(* IEC 61131-3 sources: stf-hw/web/public/sil (part 2) *)

(* HBW belt and the two RFID read points. Generated by stf-cad/hbw/sil/iec.py from the proven motion (control.py); do not edit. *)
FUNCTION_BLOCK FB_Belt
VAR_INPUT
    Enable : BOOL;        (* K0 safety relay OK AND mode = AUTO *)
    Ack : BOOL;           (* HMI acknowledge *)
    Reset : BOOL;         (* S3 reset, via the safety relay *)
    Cmd : INT;            (* job to start (0 = none), taken when READY *)
    Arg1 : INT;           (* binding: slot / bay / slot pair index *)
    I2 : BOOL;           (* phototransistor inside *)
    I3 : BOOL;           (* phototransistor outside *)
    Tag : INT;            (* the mould the record expects at RP2 *)
    ExpI2, ExpI3 : BOOL;  (* the belt's occupancy the record expects *)
    RF1_Valid, RF2_Valid : BOOL;
    RF2_Tag : INT;
END_VAR
VAR_OUTPUT
    Q1 : BOOL;           (* conveyor belt forward (M1) *)
    Q2 : BOOL;           (* conveyor belt backward (M1) *)
    Ready, Busy, Done, Fault : BOOL;   (* Done: one scan, when a job ends *)
    Alarm : INT;          (* the state whose watchdog tripped *)
    Sn : INT;             (* the active state *)
END_VAR
VAR
    Prev : INT := -1;
    Job, B1 : INT;
    Wd : TON;             (* step watchdog *)
    Tm : TON;             (* step timer *)
    WdTime : TIME;        (* the active state's watchdog; 0 = none *)
    RfSeen : BOOL;
END_VAR

(* every scan: outputs off unless the active state sets them; Done is a pulse *)
Q1 := FALSE; Q2 := FALSE; Done := FALSE;
IF NOT Enable AND Sn <> 900 THEN Sn := 900; END_IF;
Wd(IN := (Sn = Prev) AND (WdTime > T#0MS), PT := WdTime);
Tm(IN := (Sn = Prev), PT := T#1H);
IF Sn <> Prev THEN RfSeen := FALSE; END_IF;
RfSeen := RfSeen OR RF1_Valid;
Prev := Sn;
IF Wd.Q THEN Alarm := Sn; Sn := 910; END_IF;

CASE Sn OF
  0: (* INIT: power-up, all outputs off *)
      WdTime := T#0MS; IF Enable THEN Sn := 10; END_IF;
  10: (* H:check: occupancy check: I2/I3 against the record *)
      WdTime := T#0MS;
      IF (I2 = ExpI2) AND (I3 = ExpI3) THEN Sn := 100; END_IF;
  100: (* READY: homed, waiting for a job *)
      WdTime := T#0MS; Ready := TRUE; Busy := FALSE;
      IF Cmd <> 0 THEN Job := Cmd; B1 := Arg1; Busy := TRUE; Ready := FALSE;
          CASE Cmd OF 10: Sn := 1000; 12: Sn := 2000; ELSE Sn := 910; Alarm := -Cmd; END_CASE;
      END_IF;
  1000: (* belt_back.01 RP2: RP2 reads the tag of the mould going in *)
      WdTime := T#900MS;
      IF RF2_Valid AND RF2_Tag = Tag THEN Sn := 1001; END_IF;
  1001: (* belt_back.02 run->I2: belt back to the crane; RP1 reads the tag on the fly *)
      WdTime := T#8100MS;
      Q2 := TRUE;
      IF I2 AND RfSeen THEN Done := TRUE; Busy := FALSE; Sn := 100; END_IF;
  2000: (* belt_fwd.01 run->I3: belt out to the VGR hand-over; RP1 reads the tag on the fly *)
      WdTime := T#8100MS;
      Q1 := TRUE;
      IF I3 AND RfSeen THEN Sn := 2001; END_IF;
  2001: (* belt_fwd.02 RP2: RP2 reads the tag at rest and compares it with the record *)
      WdTime := T#900MS;
      IF RF2_Valid AND RF2_Tag = Tag THEN Done := TRUE; Busy := FALSE; Sn := 100; END_IF;
  900: (* ESTOP: the safety relay dropped, outputs off *)
      WdTime := T#0MS; Busy := FALSE; Ready := FALSE; IF Reset AND Enable THEN Sn := 0; END_IF;
  910: (* FAULT: a step timed out, outputs off, alarm raised *)
      WdTime := T#0MS; Fault := TRUE; Busy := FALSE; Ready := FALSE;
      IF Ack AND Enable THEN Fault := FALSE; Sn := 10; END_IF;
END_CASE;
END_FUNCTION_BLOCK

(* VGR arm and vacuum. Generated by stf-cad/hbw/sil/iec.py from the proven motion (control.py); do not edit. *)
FUNCTION_BLOCK FB_Arm
VAR_INPUT
    Enable : BOOL;        (* K0 safety relay OK AND mode = AUTO *)
    Ack : BOOL;           (* HMI acknowledge *)
    Reset : BOOL;         (* S3 reset, via the safety relay *)
    Cmd : INT;            (* job to start (0 = none), taken when READY *)
    Arg1 : INT;           (* binding: slot / bay / slot pair index *)
    I1 : BOOL;           (* reference vertical *)
    I2 : BOOL;           (* reference horizontal *)
    I3 : BOOL;           (* reference rotate *)
    I4 : BOOL;           (* vacuum switch: the cup is sealed on a part (-0.3 bar) *)
    PosPlunge : REAL;     (* plunge, from the encoder counter *)
    PosReach : REAL;     (* reach, from the encoder counter *)
    PosSwivel : REAL;     (* swivel, from the encoder counter *)
END_VAR
VAR_OUTPUT
    Q1 : BOOL;           (* vertical up (M1) *)
    Q2 : BOOL;           (* vertical down (M1) *)
    Q3 : BOOL;           (* horizontal backward (M2) *)
    Q4 : BOOL;           (* horizontal forward (M2) *)
    Q5 : BOOL;           (* rotate clockwise (M3) *)
    Q6 : BOOL;           (* rotate counter-clockwise (M3) *)
    Q8 : BOOL;           (*  *)
    Ready, Busy, Done, Fault : BOOL;   (* Done: one scan, when a job ends *)
    Alarm : INT;          (* the state whose watchdog tripped *)
    Sn : INT;             (* the active state *)
END_VAR
VAR
    Prev : INT := -1;
    Job, B1 : INT;
    Wd : TON;             (* step watchdog *)
    Tm : TON;             (* step timer *)
    WdTime : TIME;        (* the active state's watchdog; 0 = none *)
END_VAR
VAR CONSTANT
    TG_PLACE_OVEN_PLUNGE : ARRAY[1..1, 1..11] OF REAL := [240.0, 153.0, 153.0, 108.0, 104.0, 0.0, 108.0, 153.0, 153.0, 500.0, 500.0];
    TG_PLACE_OVEN_REACH : ARRAY[1..1, 1..11] OF REAL := [301.376, 365.895, 365.895, 365.895, 365.895, 0.0, 365.895, 365.895, 365.895, 0.0, 0.0];
    TG_PLACE_OVEN_SWIVEL : ARRAY[1..1, 1..11] OF REAL := [46.205, 23.396, 23.396, 23.396, 23.396, 0.0, 23.396, 23.396, 23.396, 0.0, 0.0];
    TG_BELT_TO_OVEN_PLUNGE : ARRAY[1..1, 1..10] OF REAL := [500.0, 201.0, 201.0, 156.0, 152.0, 0.0, 156.0, 201.0, 201.0, 240.0];
    TG_BELT_TO_OVEN_REACH : ARRAY[1..1, 1..10] OF REAL := [0.0, 236.857, 236.857, 236.857, 236.857, 0.0, 236.857, 236.857, 236.857, 301.376];
    TG_BELT_TO_OVEN_SWIVEL : ARRAY[1..1, 1..10] OF REAL := [0.0, 69.013, 69.013, 69.013, 69.013, 0.0, 69.013, 69.013, 69.013, 46.205];
    TG_BAY_TO_BELT_PLUNGE : ARRAY[1..3, 1..21] OF REAL := [500.0, 138.0, 138.0, 93.0, 89.0, 0.0, 93.0, 138.0, 138.0, 240.0, 240.0, 201.0, 201.0, 156.0, 152.0, 0.0, 156.0, 201.0, 201.0, 500.0, 500.0, 500.0, 138.0, 138.0, 93.0, 89.0, 0.0, 93.0, 138.0, 138.0, 240.0, 240.0, 201.0, 201.0, 156.0, 152.0, 0.0, 156.0, 201.0, 201.0, 500.0, 500.0, 500.0, 138.0, 138.0, 93.0, 89.0, 0.0, 93.0, 138.0, 138.0, 240.0, 240.0, 201.0, 201.0, 156.0, 152.0, 0.0, 156.0, 201.0, 201.0, 500.0, 500.0];
    TG_BAY_TO_BELT_REACH : ARRAY[1..3, 1..21] OF REAL := [0.0, 157.983, 157.983, 157.983, 157.983, 0.0, 157.983, 157.983, 157.983, 197.42, 197.42, 236.857, 236.857, 236.857, 236.857, 0.0, 236.857, 236.857, 236.857, 0.0, 0.0, 0.0, 155.396, 155.396, 155.396, 155.396, 0.0, 155.396, 155.396, 155.396, 196.126, 196.126, 236.857, 236.857, 236.857, 236.857, 0.0, 236.857, 236.857, 236.857, 0.0, 0.0, 0.0, 208.968, 208.968, 208.968, 208.968, 0.0, 208.968, 208.968, 208.968, 222.912, 222.912, 236.857, 236.857, 236.857, 236.857, 0.0, 236.857, 236.857, 236.857, 0.0, 0.0];
    TG_BAY_TO_BELT_SWIVEL : ARRAY[1..3, 1..21] OF REAL := [0.0, -76.518, -76.518, -76.518, -76.518, 0.0, -76.518, -76.518, -76.518, -3.752, -3.752, 69.013, 69.013, 69.013, 69.013, 0.0, 69.013, 69.013, 69.013, 0.0, 0.0, 0.0, -101.414, -101.414, -101.414, -101.414, 0.0, -101.414, -101.414, -101.414, -16.2, -16.2, 69.013, 69.013, 69.013, 69.013, 0.0, 69.013, 69.013, 69.013, 0.0, 0.0, 0.0, -122.763, -122.763, -122.763, -122.763, 0.0, -122.763, -122.763, -122.763, -26.875, -26.875, 69.013, 69.013, 69.013, 69.013, 0.0, 69.013, 69.013, 69.013, 0.0, 0.0];
    WD_BAY_TO_BELT : ARRAY[1..3, 1..21] OF TIME := [T#600MS, T#5000MS, T#600MS, T#1100MS, T#1100MS, T#1200MS, T#1100MS, T#1100MS, T#600MS, T#2300MS, T#600MS, T#2300MS, T#600MS, T#1100MS, T#1100MS, T#900MS, T#1100MS, T#1100MS, T#600MS, T#4200MS, T#600MS, T#600MS, T#5000MS, T#600MS, T#1100MS, T#1100MS, T#1200MS, T#1100MS, T#1100MS, T#600MS, T#2600MS, T#600MS, T#2600MS, T#600MS, T#1100MS, T#1100MS, T#900MS, T#1100MS, T#1100MS, T#600MS, T#4200MS, T#600MS, T#600MS, T#5000MS, T#600MS, T#1100MS, T#1100MS, T#1200MS, T#1100MS, T#1100MS, T#600MS, T#2900MS, T#600MS, T#2900MS, T#600MS, T#1100MS, T#1100MS, T#900MS, T#1100MS, T#1100MS, T#600MS, T#4200MS, T#600MS];
END_VAR

(* every scan: outputs off unless the active state sets them; Done is a pulse *)
Q1 := FALSE; Q2 := FALSE; Q3 := FALSE; Q4 := FALSE; Q5 := FALSE; Q6 := FALSE; Q8 := FALSE; Done := FALSE;
IF NOT Enable AND Sn <> 900 THEN Sn := 900; END_IF;
Wd(IN := (Sn = Prev) AND (WdTime > T#0MS), PT := WdTime);
Tm(IN := (Sn = Prev), PT := T#1H);
Prev := Sn;
IF Wd.Q THEN Alarm := Sn; Sn := 910; END_IF;

CASE Sn OF
  0: (* INIT: power-up, all outputs off *)
      WdTime := T#0MS; IF Enable THEN Sn := 10; END_IF;
  10: (* H:plunge: plunge up to the reference switch *)
      WdTime := T#6200MS;
      Q1 := TRUE;
      IF I1 THEN Sn := 11; END_IF;
  11: (* H:reach: reach back to the reference switch *)
      WdTime := T#5500MS;
      Q3 := TRUE;
      IF I2 THEN Sn := 12; END_IF;
  12: (* H:swivel: swivel to the reference switch *)
      WdTime := T#7000MS;
      Q6 := TRUE;
      IF I3 THEN Sn := 100; END_IF;
  100: (* READY: homed, waiting for a job *)
      WdTime := T#0MS; Ready := TRUE; Busy := FALSE;
      IF Cmd <> 0 THEN Job := Cmd; B1 := Arg1; Busy := TRUE; Ready := FALSE;
          CASE Cmd OF 7: Sn := 1000; 8: Sn := 2000; 9: Sn := 3000; ELSE Sn := 910; Alarm := -Cmd; END_CASE;
      END_IF;
  1000: (* place_oven.01 k11:pos: swing to the target at transit height *)
      WdTime := T#600MS;
      Q8 := TRUE;
      CASE Drive(PosPlunge, TG_PLACE_OVEN_PLUNGE[B1, 1], 0.3) OF -1: Q2 := TRUE; 1: Q1 := TRUE; END_CASE;
      CASE Drive(PosReach, TG_PLACE_OVEN_REACH[B1, 1], 0.3) OF -1: Q3 := TRUE; 1: Q4 := TRUE; END_CASE;
      CASE Drive(PosSwivel, TG_PLACE_OVEN_SWIVEL[B1, 1], 0.15) OF -1: Q6 := TRUE; 1: Q5 := TRUE; END_CASE;
      IF ABS(PosPlunge - TG_PLACE_OVEN_PLUNGE[B1, 1]) <= 4.0 AND ABS(PosReach - TG_PLACE_OVEN_REACH[B1, 1]) <= 2.5 AND ABS(PosSwivel - TG_PLACE_OVEN_SWIVEL[B1, 1]) <= 0.252 THEN Sn := 1001; END_IF;
  1001: (* place_oven.02 k12:pos: descend beside the target *)
      WdTime := T#1600MS;
      Q8 := TRUE;
      CASE Drive(PosPlunge, TG_PLACE_OVEN_PLUNGE[B1, 2], 0.3) OF -1: Q2 := TRUE; 1: Q1 := TRUE; END_CASE;
      CASE Drive(PosReach, TG_PLACE_OVEN_REACH[B1, 2], 0.3) OF -1: Q3 := TRUE; 1: Q4 := TRUE; END_CASE;
      CASE Drive(PosSwivel, TG_PLACE_OVEN_SWIVEL[B1, 2], 0.15) OF -1: Q6 := TRUE; 1: Q5 := TRUE; END_CASE;
      IF ABS(PosPlunge - TG_PLACE_OVEN_PLUNGE[B1, 2]) <= 4.0 AND ABS(PosReach - TG_PLACE_OVEN_REACH[B1, 2]) <= 2.5 AND ABS(PosSwivel - TG_PLACE_OVEN_SWIVEL[B1, 2]) <= 0.252 THEN Sn := 1002; END_IF;
  1002: (* place_oven.03 k13:pos: extend over the target *)
      WdTime := T#600MS;
      Q8 := TRUE;
      CASE Drive(PosPlunge, TG_PLACE_OVEN_PLUNGE[B1, 3], 0.3) OF -1: Q2 := TRUE; 1: Q1 := TRUE; END_CASE;
      CASE Drive(PosReach, TG_PLACE_OVEN_REACH[B1, 3], 0.3) OF -1: Q3 := TRUE; 1: Q4 := TRUE; END_CASE;
      CASE Drive(PosSwivel, TG_PLACE_OVEN_SWIVEL[B1, 3], 0.15) OF -1: Q6 := TRUE; 1: Q5 := TRUE; END_CASE;
      IF ABS(PosPlunge - TG_PLACE_OVEN_PLUNGE[B1, 3]) <= 4.0 AND ABS(PosReach - TG_PLACE_OVEN_REACH[B1, 3]) <= 2.5 AND ABS(PosSwivel - TG_PLACE_OVEN_SWIVEL[B1, 3]) <= 0.252 THEN Sn := 1003; END_IF;
  1003: (* place_oven.04 k14:pos: cup meets the cookie's top face *)
      WdTime := T#1100MS;
      Q8 := TRUE;
      CASE Drive(PosPlunge, TG_PLACE_OVEN_PLUNGE[B1, 4], 0.3) OF -1: Q2 := TRUE; 1: Q1 := TRUE; END_CASE;
      CASE Drive(PosReach, TG_PLACE_OVEN_REACH[B1, 4], 0.3) OF -1: Q3 := TRUE; 1: Q4 := TRUE; END_CASE;
      CASE Drive(PosSwivel, TG_PLACE_OVEN_SWIVEL[B1, 4], 0.15) OF -1: Q6 := TRUE; 1: Q5 := TRUE; END_CASE;
      IF ABS(PosPlunge - TG_PLACE_OVEN_PLUNGE[B1, 4]) <= 4.0 AND ABS(PosReach - TG_PLACE_OVEN_REACH[B1, 4]) <= 2.5 AND ABS(PosSwivel - TG_PLACE_OVEN_SWIVEL[B1, 4]) <= 0.252 THEN Sn := 1004; END_IF;
  1004: (* place_oven.05 k15:pos: press: the spring stem takes up the over-travel *)
      WdTime := T#1100MS;
      Q8 := TRUE;
      CASE Drive(PosPlunge, TG_PLACE_OVEN_PLUNGE[B1, 5], 0.3) OF -1: Q2 := TRUE; 1: Q1 := TRUE; END_CASE;
      CASE Drive(PosReach, TG_PLACE_OVEN_REACH[B1, 5], 0.3) OF -1: Q3 := TRUE; 1: Q4 := TRUE; END_CASE;
      CASE Drive(PosSwivel, TG_PLACE_OVEN_SWIVEL[B1, 5], 0.15) OF -1: Q6 := TRUE; 1: Q5 := TRUE; END_CASE;
      IF ABS(PosPlunge - TG_PLACE_OVEN_PLUNGE[B1, 5]) <= 4.0 AND ABS(PosReach - TG_PLACE_OVEN_REACH[B1, 5]) <= 2.5 AND ABS(PosSwivel - TG_PLACE_OVEN_SWIVEL[B1, 5]) <= 0.252 THEN Sn := 1005; END_IF;
  1005: (* place_oven.06 k16:vac: Q8 off: the cookie is released (I4 drops) *)
      WdTime := T#900MS;
      IF NOT I4 THEN Sn := 1006; END_IF;
  1006: (* place_oven.07 k17:pos: spring relaxes *)
      WdTime := T#1100MS;
      CASE Drive(PosPlunge, TG_PLACE_OVEN_PLUNGE[B1, 7], 0.3) OF -1: Q2 := TRUE; 1: Q1 := TRUE; END_CASE;
      CASE Drive(PosReach, TG_PLACE_OVEN_REACH[B1, 7], 0.3) OF -1: Q3 := TRUE; 1: Q4 := TRUE; END_CASE;
      CASE Drive(PosSwivel, TG_PLACE_OVEN_SWIVEL[B1, 7], 0.15) OF -1: Q6 := TRUE; 1: Q5 := TRUE; END_CASE;
      IF ABS(PosPlunge - TG_PLACE_OVEN_PLUNGE[B1, 7]) <= 4.0 AND ABS(PosReach - TG_PLACE_OVEN_REACH[B1, 7]) <= 2.5 AND ABS(PosSwivel - TG_PLACE_OVEN_SWIVEL[B1, 7]) <= 0.252 THEN Sn := 1007; END_IF;
  1007: (* place_oven.08 k18:pos: lift clear *)
      WdTime := T#1100MS;
      CASE Drive(PosPlunge, TG_PLACE_OVEN_PLUNGE[B1, 8], 0.3) OF -1: Q2 := TRUE; 1: Q1 := TRUE; END_CASE;
      CASE Drive(PosReach, TG_PLACE_OVEN_REACH[B1, 8], 0.3) OF -1: Q3 := TRUE; 1: Q4 := TRUE; END_CASE;
      CASE Drive(PosSwivel, TG_PLACE_OVEN_SWIVEL[B1, 8], 0.15) OF -1: Q6 := TRUE; 1: Q5 := TRUE; END_CASE;
      IF ABS(PosPlunge - TG_PLACE_OVEN_PLUNGE[B1, 8]) <= 4.0 AND ABS(PosReach - TG_PLACE_OVEN_REACH[B1, 8]) <= 2.5 AND ABS(PosSwivel - TG_PLACE_OVEN_SWIVEL[B1, 8]) <= 0.252 THEN Sn := 1008; END_IF;
  1008: (* place_oven.09 k19:pos: retract out from the station *)
      WdTime := T#600MS;
      CASE Drive(PosPlunge, TG_PLACE_OVEN_PLUNGE[B1, 9], 0.3) OF -1: Q2 := TRUE; 1: Q1 := TRUE; END_CASE;
      CASE Drive(PosReach, TG_PLACE_OVEN_REACH[B1, 9], 0.3) OF -1: Q3 := TRUE; 1: Q4 := TRUE; END_CASE;
      CASE Drive(PosSwivel, TG_PLACE_OVEN_SWIVEL[B1, 9], 0.15) OF -1: Q6 := TRUE; 1: Q5 := TRUE; END_CASE;
      IF ABS(PosPlunge - TG_PLACE_OVEN_PLUNGE[B1, 9]) <= 4.0 AND ABS(PosReach - TG_PLACE_OVEN_REACH[B1, 9]) <= 2.5 AND ABS(PosSwivel - TG_PLACE_OVEN_SWIVEL[B1, 9]) <= 0.252 THEN Sn := 1009; END_IF;
  1009: (* place_oven.10 k20:pos: rise to transit height *)
      WdTime := T#5100MS;
      CASE Drive(PosPlunge, TG_PLACE_OVEN_PLUNGE[B1, 10], 0.3) OF -1: Q2 := TRUE; 1: Q1 := TRUE; END_CASE;
      CASE Drive(PosReach, TG_PLACE_OVEN_REACH[B1, 10], 0.3) OF -1: Q3 := TRUE; 1: Q4 := TRUE; END_CASE;
      CASE Drive(PosSwivel, TG_PLACE_OVEN_SWIVEL[B1, 10], 0.15) OF -1: Q6 := TRUE; 1: Q5 := TRUE; END_CASE;
      IF ABS(PosPlunge - TG_PLACE_OVEN_PLUNGE[B1, 10]) <= 4.0 AND ABS(PosReach - TG_PLACE_OVEN_REACH[B1, 10]) <= 2.5 AND ABS(PosSwivel - TG_PLACE_OVEN_SWIVEL[B1, 10]) <= 0.252 THEN Sn := 1010; END_IF;
  1010: (* place_oven.11 k21:pos: VGR back home *)
      WdTime := T#600MS;
      CASE Drive(PosPlunge, TG_PLACE_OVEN_PLUNGE[B1, 11], 0.3) OF -1: Q2 := TRUE; 1: Q1 := TRUE; END_CASE;
      CASE Drive(PosReach, TG_PLACE_OVEN_REACH[B1, 11], 0.3) OF -1: Q3 := TRUE; 1: Q4 := TRUE; END_CASE;
      CASE Drive(PosSwivel, TG_PLACE_OVEN_SWIVEL[B1, 11], 0.15) OF -1: Q6 := TRUE; 1: Q5 := TRUE; END_CASE;
      IF ABS(PosPlunge - TG_PLACE_OVEN_PLUNGE[B1, 11]) <= 4.0 AND ABS(PosReach - TG_PLACE_OVEN_REACH[B1, 11]) <= 2.5 AND ABS(PosSwivel - TG_PLACE_OVEN_SWIVEL[B1, 11]) <= 0.252 THEN Done := TRUE; Busy := FALSE; Sn := 100; END_IF;
  2000: (* belt_to_oven.01 k1:pos: swing to the source at transit height *)
      WdTime := T#600MS;
      CASE Drive(PosPlunge, TG_BELT_TO_OVEN_PLUNGE[B1, 1], 0.3) OF -1: Q2 := TRUE; 1: Q1 := TRUE; END_CASE;
      CASE Drive(PosReach, TG_BELT_TO_OVEN_REACH[B1, 1], 0.3) OF -1: Q3 := TRUE; 1: Q4 := TRUE; END_CASE;
      CASE Drive(PosSwivel, TG_BELT_TO_OVEN_SWIVEL[B1, 1], 0.15) OF -1: Q6 := TRUE; 1: Q5 := TRUE; END_CASE;
      IF ABS(PosPlunge - TG_BELT_TO_OVEN_PLUNGE[B1, 1]) <= 4.0 AND ABS(PosReach - TG_BELT_TO_OVEN_REACH[B1, 1]) <= 2.5 AND ABS(PosSwivel - TG_BELT_TO_OVEN_SWIVEL[B1, 1]) <= 0.252 THEN Sn := 2001; END_IF;
  2001: (* belt_to_oven.02 k2:pos: descend beside the source *)
      WdTime := T#4200MS;
      CASE Drive(PosPlunge, TG_BELT_TO_OVEN_PLUNGE[B1, 2], 0.3) OF -1: Q2 := TRUE; 1: Q1 := TRUE; END_CASE;
      CASE Drive(PosReach, TG_BELT_TO_OVEN_REACH[B1, 2], 0.3) OF -1: Q3 := TRUE; 1: Q4 := TRUE; END_CASE;
      CASE Drive(PosSwivel, TG_BELT_TO_OVEN_SWIVEL[B1, 2], 0.15) OF -1: Q6 := TRUE; 1: Q5 := TRUE; END_CASE;
      IF ABS(PosPlunge - TG_BELT_TO_OVEN_PLUNGE[B1, 2]) <= 4.0 AND ABS(PosReach - TG_BELT_TO_OVEN_REACH[B1, 2]) <= 2.5 AND ABS(PosSwivel - TG_BELT_TO_OVEN_SWIVEL[B1, 2]) <= 0.252 THEN Sn := 2002; END_IF;
  2002: (* belt_to_oven.03 k3:pos: extend over the source *)
      WdTime := T#600MS;
      CASE Drive(PosPlunge, TG_BELT_TO_OVEN_PLUNGE[B1, 3], 0.3) OF -1: Q2 := TRUE; 1: Q1 := TRUE; END_CASE;
      CASE Drive(PosReach, TG_BELT_TO_OVEN_REACH[B1, 3], 0.3) OF -1: Q3 := TRUE; 1: Q4 := TRUE; END_CASE;
      CASE Drive(PosSwivel, TG_BELT_TO_OVEN_SWIVEL[B1, 3], 0.15) OF -1: Q6 := TRUE; 1: Q5 := TRUE; END_CASE;
      IF ABS(PosPlunge - TG_BELT_TO_OVEN_PLUNGE[B1, 3]) <= 4.0 AND ABS(PosReach - TG_BELT_TO_OVEN_REACH[B1, 3]) <= 2.5 AND ABS(PosSwivel - TG_BELT_TO_OVEN_SWIVEL[B1, 3]) <= 0.252 THEN Sn := 2003; END_IF;
  2003: (* belt_to_oven.04 k4:pos: cup meets the cookie's top face *)
      WdTime := T#1100MS;
      CASE Drive(PosPlunge, TG_BELT_TO_OVEN_PLUNGE[B1, 4], 0.3) OF -1: Q2 := TRUE; 1: Q1 := TRUE; END_CASE;
      CASE Drive(PosReach, TG_BELT_TO_OVEN_REACH[B1, 4], 0.3) OF -1: Q3 := TRUE; 1: Q4 := TRUE; END_CASE;
      CASE Drive(PosSwivel, TG_BELT_TO_OVEN_SWIVEL[B1, 4], 0.15) OF -1: Q6 := TRUE; 1: Q5 := TRUE; END_CASE;
      IF ABS(PosPlunge - TG_BELT_TO_OVEN_PLUNGE[B1, 4]) <= 4.0 AND ABS(PosReach - TG_BELT_TO_OVEN_REACH[B1, 4]) <= 2.5 AND ABS(PosSwivel - TG_BELT_TO_OVEN_SWIVEL[B1, 4]) <= 0.252 THEN Sn := 2004; END_IF;
  2004: (* belt_to_oven.05 k5:pos: press: the spring stem takes up the over-travel *)
      WdTime := T#1100MS;
      CASE Drive(PosPlunge, TG_BELT_TO_OVEN_PLUNGE[B1, 5], 0.3) OF -1: Q2 := TRUE; 1: Q1 := TRUE; END_CASE;
      CASE Drive(PosReach, TG_BELT_TO_OVEN_REACH[B1, 5], 0.3) OF -1: Q3 := TRUE; 1: Q4 := TRUE; END_CASE;
      CASE Drive(PosSwivel, TG_BELT_TO_OVEN_SWIVEL[B1, 5], 0.15) OF -1: Q6 := TRUE; 1: Q5 := TRUE; END_CASE;
      IF ABS(PosPlunge - TG_BELT_TO_OVEN_PLUNGE[B1, 5]) <= 4.0 AND ABS(PosReach - TG_BELT_TO_OVEN_REACH[B1, 5]) <= 2.5 AND ABS(PosSwivel - TG_BELT_TO_OVEN_SWIVEL[B1, 5]) <= 0.252 THEN Sn := 2005; END_IF;
  2005: (* belt_to_oven.06 k6:vac: Q8 vacuum on: the cup seals on the cookie (I4 made) *)
      WdTime := T#1200MS;
      Q8 := TRUE;
      IF I4 THEN Sn := 2006; END_IF;
  2006: (* belt_to_oven.07 k7:pos: spring relaxes - seal holds *)
      WdTime := T#1100MS;
      Q8 := TRUE;
      CASE Drive(PosPlunge, TG_BELT_TO_OVEN_PLUNGE[B1, 7], 0.3) OF -1: Q2 := TRUE; 1: Q1 := TRUE; END_CASE;
      CASE Drive(PosReach, TG_BELT_TO_OVEN_REACH[B1, 7], 0.3) OF -1: Q3 := TRUE; 1: Q4 := TRUE; END_CASE;
      CASE Drive(PosSwivel, TG_BELT_TO_OVEN_SWIVEL[B1, 7], 0.15) OF -1: Q6 := TRUE; 1: Q5 := TRUE; END_CASE;
      IF ABS(PosPlunge - TG_BELT_TO_OVEN_PLUNGE[B1, 7]) <= 4.0 AND ABS(PosReach - TG_BELT_TO_OVEN_REACH[B1, 7]) <= 2.5 AND ABS(PosSwivel - TG_BELT_TO_OVEN_SWIVEL[B1, 7]) <= 0.252 THEN Sn := 2007; END_IF;
  2007: (* belt_to_oven.08 k8:pos: lift the cookie clear *)
      WdTime := T#1100MS;
      Q8 := TRUE;
      CASE Drive(PosPlunge, TG_BELT_TO_OVEN_PLUNGE[B1, 8], 0.3) OF -1: Q2 := TRUE; 1: Q1 := TRUE; END_CASE;
      CASE Drive(PosReach, TG_BELT_TO_OVEN_REACH[B1, 8], 0.3) OF -1: Q3 := TRUE; 1: Q4 := TRUE; END_CASE;
      CASE Drive(PosSwivel, TG_BELT_TO_OVEN_SWIVEL[B1, 8], 0.15) OF -1: Q6 := TRUE; 1: Q5 := TRUE; END_CASE;
      IF ABS(PosPlunge - TG_BELT_TO_OVEN_PLUNGE[B1, 8]) <= 4.0 AND ABS(PosReach - TG_BELT_TO_OVEN_REACH[B1, 8]) <= 2.5 AND ABS(PosSwivel - TG_BELT_TO_OVEN_SWIVEL[B1, 8]) <= 0.252 THEN Sn := 2008; END_IF;
  2008: (* belt_to_oven.09 k9:pos: retract out from the station *)
      WdTime := T#600MS;
      Q8 := TRUE;
      CASE Drive(PosPlunge, TG_BELT_TO_OVEN_PLUNGE[B1, 9], 0.3) OF -1: Q2 := TRUE; 1: Q1 := TRUE; END_CASE;
      CASE Drive(PosReach, TG_BELT_TO_OVEN_REACH[B1, 9], 0.3) OF -1: Q3 := TRUE; 1: Q4 := TRUE; END_CASE;
      CASE Drive(PosSwivel, TG_BELT_TO_OVEN_SWIVEL[B1, 9], 0.15) OF -1: Q6 := TRUE; 1: Q5 := TRUE; END_CASE;
      IF ABS(PosPlunge - TG_BELT_TO_OVEN_PLUNGE[B1, 9]) <= 4.0 AND ABS(PosReach - TG_BELT_TO_OVEN_REACH[B1, 9]) <= 2.5 AND ABS(PosSwivel - TG_BELT_TO_OVEN_SWIVEL[B1, 9]) <= 0.252 THEN Sn := 2009; END_IF;
  2009: (* belt_to_oven.10 k10:pos: rise to transit height *)
      WdTime := T#1300MS;
      Q8 := TRUE;
      CASE Drive(PosPlunge, TG_BELT_TO_OVEN_PLUNGE[B1, 10], 0.3) OF -1: Q2 := TRUE; 1: Q1 := TRUE; END_CASE;
      CASE Drive(PosReach, TG_BELT_TO_OVEN_REACH[B1, 10], 0.3) OF -1: Q3 := TRUE; 1: Q4 := TRUE; END_CASE;
      CASE Drive(PosSwivel, TG_BELT_TO_OVEN_SWIVEL[B1, 10], 0.15) OF -1: Q6 := TRUE; 1: Q5 := TRUE; END_CASE;
      IF ABS(PosPlunge - TG_BELT_TO_OVEN_PLUNGE[B1, 10]) <= 4.0 AND ABS(PosReach - TG_BELT_TO_OVEN_REACH[B1, 10]) <= 2.5 AND ABS(PosSwivel - TG_BELT_TO_OVEN_SWIVEL[B1, 10]) <= 0.252 THEN Done := TRUE; Busy := FALSE; Sn := 100; END_IF;
  3000: (* bay_to_belt.01 k1:pos: swing to the source at transit height *)
      WdTime := T#600MS;
      CASE Drive(PosPlunge, TG_BAY_TO_BELT_PLUNGE[B1, 1], 0.3) OF -1: Q2 := TRUE; 1: Q1 := TRUE; END_CASE;
      CASE Drive(PosReach, TG_BAY_TO_BELT_REACH[B1, 1], 0.3) OF -1: Q3 := TRUE; 1: Q4 := TRUE; END_CASE;
      CASE Drive(PosSwivel, TG_BAY_TO_BELT_SWIVEL[B1, 1], 0.15) OF -1: Q6 := TRUE; 1: Q5 := TRUE; END_CASE;
      IF ABS(PosPlunge - TG_BAY_TO_BELT_PLUNGE[B1, 1]) <= 4.0 AND ABS(PosReach - TG_BAY_TO_BELT_REACH[B1, 1]) <= 2.5 AND ABS(PosSwivel - TG_BAY_TO_BELT_SWIVEL[B1, 1]) <= 0.252 THEN Sn := 3001; END_IF;
  3001: (* bay_to_belt.02 k2:pos: descend beside the source *)
      WdTime := T#5000MS;
      CASE Drive(PosPlunge, TG_BAY_TO_BELT_PLUNGE[B1, 2], 0.3) OF -1: Q2 := TRUE; 1: Q1 := TRUE; END_CASE;
      CASE Drive(PosReach, TG_BAY_TO_BELT_REACH[B1, 2], 0.3) OF -1: Q3 := TRUE; 1: Q4 := TRUE; END_CASE;
      CASE Drive(PosSwivel, TG_BAY_TO_BELT_SWIVEL[B1, 2], 0.15) OF -1: Q6 := TRUE; 1: Q5 := TRUE; END_CASE;
      IF ABS(PosPlunge - TG_BAY_TO_BELT_PLUNGE[B1, 2]) <= 4.0 AND ABS(PosReach - TG_BAY_TO_BELT_REACH[B1, 2]) <= 2.5 AND ABS(PosSwivel - TG_BAY_TO_BELT_SWIVEL[B1, 2]) <= 0.252 THEN Sn := 3002; END_IF;
  3002: (* bay_to_belt.03 k3:pos: extend over the source *)
      WdTime := T#600MS;
      CASE Drive(PosPlunge, TG_BAY_TO_BELT_PLUNGE[B1, 3], 0.3) OF -1: Q2 := TRUE; 1: Q1 := TRUE; END_CASE;
      CASE Drive(PosReach, TG_BAY_TO_BELT_REACH[B1, 3], 0.3) OF -1: Q3 := TRUE; 1: Q4 := TRUE; END_CASE;
      CASE Drive(PosSwivel, TG_BAY_TO_BELT_SWIVEL[B1, 3], 0.15) OF -1: Q6 := TRUE; 1: Q5 := TRUE; END_CASE;
      IF ABS(PosPlunge - TG_BAY_TO_BELT_PLUNGE[B1, 3]) <= 4.0 AND ABS(PosReach - TG_BAY_TO_BELT_REACH[B1, 3]) <= 2.5 AND ABS(PosSwivel - TG_BAY_TO_BELT_SWIVEL[B1, 3]) <= 0.252 THEN Sn := 3003; END_IF;
  3003: (* bay_to_belt.04 k4:pos: cup meets the cookie's top face *)
      WdTime := T#1100MS;
      CASE Drive(PosPlunge, TG_BAY_TO_BELT_PLUNGE[B1, 4], 0.3) OF -1: Q2 := TRUE; 1: Q1 := TRUE; END_CASE;
      CASE Drive(PosReach, TG_BAY_TO_BELT_REACH[B1, 4], 0.3) OF -1: Q3 := TRUE; 1: Q4 := TRUE; END_CASE;
      CASE Drive(PosSwivel, TG_BAY_TO_BELT_SWIVEL[B1, 4], 0.15) OF -1: Q6 := TRUE; 1: Q5 := TRUE; END_CASE;
      IF ABS(PosPlunge - TG_BAY_TO_BELT_PLUNGE[B1, 4]) <= 4.0 AND ABS(PosReach - TG_BAY_TO_BELT_REACH[B1, 4]) <= 2.5 AND ABS(PosSwivel - TG_BAY_TO_BELT_SWIVEL[B1, 4]) <= 0.252 THEN Sn := 3004; END_IF;
  3004: (* bay_to_belt.05 k5:pos: press: the spring stem takes up the over-travel *)
      WdTime := T#1100MS;
      CASE Drive(PosPlunge, TG_BAY_TO_BELT_PLUNGE[B1, 5], 0.3) OF -1: Q2 := TRUE; 1: Q1 := TRUE; END_CASE;
      CASE Drive(PosReach, TG_BAY_TO_BELT_REACH[B1, 5], 0.3) OF -1: Q3 := TRUE; 1: Q4 := TRUE; END_CASE;
      CASE Drive(PosSwivel, TG_BAY_TO_BELT_SWIVEL[B1, 5], 0.15) OF -1: Q6 := TRUE; 1: Q5 := TRUE; END_CASE;
      IF ABS(PosPlunge - TG_BAY_TO_BELT_PLUNGE[B1, 5]) <= 4.0 AND ABS(PosReach - TG_BAY_TO_BELT_REACH[B1, 5]) <= 2.5 AND ABS(PosSwivel - TG_BAY_TO_BELT_SWIVEL[B1, 5]) <= 0.252 THEN Sn := 3005; END_IF;
  3005: (* bay_to_belt.06 k6:vac: Q8 vacuum on: the cup seals on the cookie (I4 made) *)
      WdTime := T#1200MS;
      Q8 := TRUE;
      IF I4 THEN Sn := 3006; END_IF;
  3006: (* bay_to_belt.07 k7:pos: spring relaxes - seal holds *)
      WdTime := T#1100MS;
      Q8 := TRUE;
      CASE Drive(PosPlunge, TG_BAY_TO_BELT_PLUNGE[B1, 7], 0.3) OF -1: Q2 := TRUE; 1: Q1 := TRUE; END_CASE;
      CASE Drive(PosReach, TG_BAY_TO_BELT_REACH[B1, 7], 0.3) OF -1: Q3 := TRUE; 1: Q4 := TRUE; END_CASE;
      CASE Drive(PosSwivel, TG_BAY_TO_BELT_SWIVEL[B1, 7], 0.15) OF -1: Q6 := TRUE; 1: Q5 := TRUE; END_CASE;
      IF ABS(PosPlunge - TG_BAY_TO_BELT_PLUNGE[B1, 7]) <= 4.0 AND ABS(PosReach - TG_BAY_TO_BELT_REACH[B1, 7]) <= 2.5 AND ABS(PosSwivel - TG_BAY_TO_BELT_SWIVEL[B1, 7]) <= 0.252 THEN Sn := 3007; END_IF;
  3007: (* bay_to_belt.08 k8:pos: lift the cookie clear *)
      WdTime := T#1100MS;
      Q8 := TRUE;
      CASE Drive(PosPlunge, TG_BAY_TO_BELT_PLUNGE[B1, 8], 0.3) OF -1: Q2 := TRUE; 1: Q1 := TRUE; END_CASE;
      CASE Drive(PosReach, TG_BAY_TO_BELT_REACH[B1, 8], 0.3) OF -1: Q3 := TRUE; 1: Q4 := TRUE; END_CASE;
      CASE Drive(PosSwivel, TG_BAY_TO_BELT_SWIVEL[B1, 8], 0.15) OF -1: Q6 := TRUE; 1: Q5 := TRUE; END_CASE;
      IF ABS(PosPlunge - TG_BAY_TO_BELT_PLUNGE[B1, 8]) <= 4.0 AND ABS(PosReach - TG_BAY_TO_BELT_REACH[B1, 8]) <= 2.5 AND ABS(PosSwivel - TG_BAY_TO_BELT_SWIVEL[B1, 8]) <= 0.252 THEN Sn := 3008; END_IF;
  3008: (* bay_to_belt.09 k9:pos: retract out from the station *)
      WdTime := T#600MS;
      Q8 := TRUE;
      CASE Drive(PosPlunge, TG_BAY_TO_BELT_PLUNGE[B1, 9], 0.3) OF -1: Q2 := TRUE; 1: Q1 := TRUE; END_CASE;
      CASE Drive(PosReach, TG_BAY_TO_BELT_REACH[B1, 9], 0.3) OF -1: Q3 := TRUE; 1: Q4 := TRUE; END_CASE;
      CASE Drive(PosSwivel, TG_BAY_TO_BELT_SWIVEL[B1, 9], 0.15) OF -1: Q6 := TRUE; 1: Q5 := TRUE; END_CASE;
      IF ABS(PosPlunge - TG_BAY_TO_BELT_PLUNGE[B1, 9]) <= 4.0 AND ABS(PosReach - TG_BAY_TO_BELT_REACH[B1, 9]) <= 2.5 AND ABS(PosSwivel - TG_BAY_TO_BELT_SWIVEL[B1, 9]) <= 0.252 THEN Sn := 3009; END_IF;
  3009: (* bay_to_belt.10 k10:pos: rise to transit height *)
      WdTime := WD_BAY_TO_BELT[B1, 10];
      Q8 := TRUE;
      CASE Drive(PosPlunge, TG_BAY_TO_BELT_PLUNGE[B1, 10], 0.3) OF -1: Q2 := TRUE; 1: Q1 := TRUE; END_CASE;
      CASE Drive(PosReach, TG_BAY_TO_BELT_REACH[B1, 10], 0.3) OF -1: Q3 := TRUE; 1: Q4 := TRUE; END_CASE;
      CASE Drive(PosSwivel, TG_BAY_TO_BELT_SWIVEL[B1, 10], 0.15) OF -1: Q6 := TRUE; 1: Q5 := TRUE; END_CASE;
      IF ABS(PosPlunge - TG_BAY_TO_BELT_PLUNGE[B1, 10]) <= 4.0 AND ABS(PosReach - TG_BAY_TO_BELT_REACH[B1, 10]) <= 2.5 AND ABS(PosSwivel - TG_BAY_TO_BELT_SWIVEL[B1, 10]) <= 0.252 THEN Sn := 3010; END_IF;
  3010: (* bay_to_belt.11 k11:pos: swing to the target at transit height *)
      WdTime := T#600MS;
      Q8 := TRUE;
      CASE Drive(PosPlunge, TG_BAY_TO_BELT_PLUNGE[B1, 11], 0.3) OF -1: Q2 := TRUE; 1: Q1 := TRUE; END_CASE;
      CASE Drive(PosReach, TG_BAY_TO_BELT_REACH[B1, 11], 0.3) OF -1: Q3 := TRUE; 1: Q4 := TRUE; END_CASE;
      CASE Drive(PosSwivel, TG_BAY_TO_BELT_SWIVEL[B1, 11], 0.15) OF -1: Q6 := TRUE; 1: Q5 := TRUE; END_CASE;
      IF ABS(PosPlunge - TG_BAY_TO_BELT_PLUNGE[B1, 11]) <= 4.0 AND ABS(PosReach - TG_BAY_TO_BELT_REACH[B1, 11]) <= 2.5 AND ABS(PosSwivel - TG_BAY_TO_BELT_SWIVEL[B1, 11]) <= 0.252 THEN Sn := 3011; END_IF;
  3011: (* bay_to_belt.12 k12:pos: descend beside the target *)
      WdTime := WD_BAY_TO_BELT[B1, 12];
      Q8 := TRUE;
      CASE Drive(PosPlunge, TG_BAY_TO_BELT_PLUNGE[B1, 12], 0.3) OF -1: Q2 := TRUE; 1: Q1 := TRUE; END_CASE;
      CASE Drive(PosReach, TG_BAY_TO_BELT_REACH[B1, 12], 0.3) OF -1: Q3 := TRUE; 1: Q4 := TRUE; END_CASE;
      CASE Drive(PosSwivel, TG_BAY_TO_BELT_SWIVEL[B1, 12], 0.15) OF -1: Q6 := TRUE; 1: Q5 := TRUE; END_CASE;
      IF ABS(PosPlunge - TG_BAY_TO_BELT_PLUNGE[B1, 12]) <= 4.0 AND ABS(PosReach - TG_BAY_TO_BELT_REACH[B1, 12]) <= 2.5 AND ABS(PosSwivel - TG_BAY_TO_BELT_SWIVEL[B1, 12]) <= 0.252 THEN Sn := 3012; END_IF;
  3012: (* bay_to_belt.13 k13:pos: extend over the target *)
      WdTime := T#600MS;
      Q8 := TRUE;
      CASE Drive(PosPlunge, TG_BAY_TO_BELT_PLUNGE[B1, 13], 0.3) OF -1: Q2 := TRUE; 1: Q1 := TRUE; END_CASE;
      CASE Drive(PosReach, TG_BAY_TO_BELT_REACH[B1, 13], 0.3) OF -1: Q3 := TRUE; 1: Q4 := TRUE; END_CASE;
      CASE Drive(PosSwivel, TG_BAY_TO_BELT_SWIVEL[B1, 13], 0.15) OF -1: Q6 := TRUE; 1: Q5 := TRUE; END_CASE;
      IF ABS(PosPlunge - TG_BAY_TO_BELT_PLUNGE[B1, 13]) <= 4.0 AND ABS(PosReach - TG_BAY_TO_BELT_REACH[B1, 13]) <= 2.5 AND ABS(PosSwivel - TG_BAY_TO_BELT_SWIVEL[B1, 13]) <= 0.252 THEN Sn := 3013; END_IF;
  3013: (* bay_to_belt.14 k14:pos: cup meets the cookie's top face *)
      WdTime := T#1100MS;
      Q8 := TRUE;
      CASE Drive(PosPlunge, TG_BAY_TO_BELT_PLUNGE[B1, 14], 0.3) OF -1: Q2 := TRUE; 1: Q1 := TRUE; END_CASE;
      CASE Drive(PosReach, TG_BAY_TO_BELT_REACH[B1, 14], 0.3) OF -1: Q3 := TRUE; 1: Q4 := TRUE; END_CASE;
      CASE Drive(PosSwivel, TG_BAY_TO_BELT_SWIVEL[B1, 14], 0.15) OF -1: Q6 := TRUE; 1: Q5 := TRUE; END_CASE;
      IF ABS(PosPlunge - TG_BAY_TO_BELT_PLUNGE[B1, 14]) <= 4.0 AND ABS(PosReach - TG_BAY_TO_BELT_REACH[B1, 14]) <= 2.5 AND ABS(PosSwivel - TG_BAY_TO_BELT_SWIVEL[B1, 14]) <= 0.252 THEN Sn := 3014; END_IF;
  3014: (* bay_to_belt.15 k15:pos: press: the spring stem takes up the over-travel *)
      WdTime := T#1100MS;
      Q8 := TRUE;
      CASE Drive(PosPlunge, TG_BAY_TO_BELT_PLUNGE[B1, 15], 0.3) OF -1: Q2 := TRUE; 1: Q1 := TRUE; END_CASE;
      CASE Drive(PosReach, TG_BAY_TO_BELT_REACH[B1, 15], 0.3) OF -1: Q3 := TRUE; 1: Q4 := TRUE; END_CASE;
      CASE Drive(PosSwivel, TG_BAY_TO_BELT_SWIVEL[B1, 15], 0.15) OF -1: Q6 := TRUE; 1: Q5 := TRUE; END_CASE;
      IF ABS(PosPlunge - TG_BAY_TO_BELT_PLUNGE[B1, 15]) <= 4.0 AND ABS(PosReach - TG_BAY_TO_BELT_REACH[B1, 15]) <= 2.5 AND ABS(PosSwivel - TG_BAY_TO_BELT_SWIVEL[B1, 15]) <= 0.252 THEN Sn := 3015; END_IF;
  3015: (* bay_to_belt.16 k16:vac: Q8 off: the cookie is released (I4 drops) *)
      WdTime := T#900MS;
      IF NOT I4 THEN Sn := 3016; END_IF;
  3016: (* bay_to_belt.17 k17:pos: spring relaxes *)
      WdTime := T#1100MS;
      CASE Drive(PosPlunge, TG_BAY_TO_BELT_PLUNGE[B1, 17], 0.3) OF -1: Q2 := TRUE; 1: Q1 := TRUE; END_CASE;
      CASE Drive(PosReach, TG_BAY_TO_BELT_REACH[B1, 17], 0.3) OF -1: Q3 := TRUE; 1: Q4 := TRUE; END_CASE;
      CASE Drive(PosSwivel, TG_BAY_TO_BELT_SWIVEL[B1, 17], 0.15) OF -1: Q6 := TRUE; 1: Q5 := TRUE; END_CASE;
      IF ABS(PosPlunge - TG_BAY_TO_BELT_PLUNGE[B1, 17]) <= 4.0 AND ABS(PosReach - TG_BAY_TO_BELT_REACH[B1, 17]) <= 2.5 AND ABS(PosSwivel - TG_BAY_TO_BELT_SWIVEL[B1, 17]) <= 0.252 THEN Sn := 3017; END_IF;
  3017: (* bay_to_belt.18 k18:pos: lift clear *)
      WdTime := T#1100MS;
      CASE Drive(PosPlunge, TG_BAY_TO_BELT_PLUNGE[B1, 18], 0.3) OF -1: Q2 := TRUE; 1: Q1 := TRUE; END_CASE;
      CASE Drive(PosReach, TG_BAY_TO_BELT_REACH[B1, 18], 0.3) OF -1: Q3 := TRUE; 1: Q4 := TRUE; END_CASE;
      CASE Drive(PosSwivel, TG_BAY_TO_BELT_SWIVEL[B1, 18], 0.15) OF -1: Q6 := TRUE; 1: Q5 := TRUE; END_CASE;
      IF ABS(PosPlunge - TG_BAY_TO_BELT_PLUNGE[B1, 18]) <= 4.0 AND ABS(PosReach - TG_BAY_TO_BELT_REACH[B1, 18]) <= 2.5 AND ABS(PosSwivel - TG_BAY_TO_BELT_SWIVEL[B1, 18]) <= 0.252 THEN Sn := 3018; END_IF;
  3018: (* bay_to_belt.19 k19:pos: retract out from the station *)
      WdTime := T#600MS;
      CASE Drive(PosPlunge, TG_BAY_TO_BELT_PLUNGE[B1, 19], 0.3) OF -1: Q2 := TRUE; 1: Q1 := TRUE; END_CASE;
      CASE Drive(PosReach, TG_BAY_TO_BELT_REACH[B1, 19], 0.3) OF -1: Q3 := TRUE; 1: Q4 := TRUE; END_CASE;
      CASE Drive(PosSwivel, TG_BAY_TO_BELT_SWIVEL[B1, 19], 0.15) OF -1: Q6 := TRUE; 1: Q5 := TRUE; END_CASE;
      IF ABS(PosPlunge - TG_BAY_TO_BELT_PLUNGE[B1, 19]) <= 4.0 AND ABS(PosReach - TG_BAY_TO_BELT_REACH[B1, 19]) <= 2.5 AND ABS(PosSwivel - TG_BAY_TO_BELT_SWIVEL[B1, 19]) <= 0.252 THEN Sn := 3019; END_IF;
  3019: (* bay_to_belt.20 k20:pos: rise to transit height *)
      WdTime := T#4200MS;
      CASE Drive(PosPlunge, TG_BAY_TO_BELT_PLUNGE[B1, 20], 0.3) OF -1: Q2 := TRUE; 1: Q1 := TRUE; END_CASE;
      CASE Drive(PosReach, TG_BAY_TO_BELT_REACH[B1, 20], 0.3) OF -1: Q3 := TRUE; 1: Q4 := TRUE; END_CASE;
      CASE Drive(PosSwivel, TG_BAY_TO_BELT_SWIVEL[B1, 20], 0.15) OF -1: Q6 := TRUE; 1: Q5 := TRUE; END_CASE;
      IF ABS(PosPlunge - TG_BAY_TO_BELT_PLUNGE[B1, 20]) <= 4.0 AND ABS(PosReach - TG_BAY_TO_BELT_REACH[B1, 20]) <= 2.5 AND ABS(PosSwivel - TG_BAY_TO_BELT_SWIVEL[B1, 20]) <= 0.252 THEN Sn := 3020; END_IF;
  3020: (* bay_to_belt.21 k21:pos: VGR back home *)
      WdTime := T#600MS;
      CASE Drive(PosPlunge, TG_BAY_TO_BELT_PLUNGE[B1, 21], 0.3) OF -1: Q2 := TRUE; 1: Q1 := TRUE; END_CASE;
      CASE Drive(PosReach, TG_BAY_TO_BELT_REACH[B1, 21], 0.3) OF -1: Q3 := TRUE; 1: Q4 := TRUE; END_CASE;
      CASE Drive(PosSwivel, TG_BAY_TO_BELT_SWIVEL[B1, 21], 0.15) OF -1: Q6 := TRUE; 1: Q5 := TRUE; END_CASE;
      IF ABS(PosPlunge - TG_BAY_TO_BELT_PLUNGE[B1, 21]) <= 4.0 AND ABS(PosReach - TG_BAY_TO_BELT_REACH[B1, 21]) <= 2.5 AND ABS(PosSwivel - TG_BAY_TO_BELT_SWIVEL[B1, 21]) <= 0.252 THEN Done := TRUE; Busy := FALSE; Sn := 100; END_IF;
  900: (* ESTOP: the safety relay dropped, outputs off *)
      WdTime := T#0MS; Busy := FALSE; Ready := FALSE; IF Reset AND Enable THEN Sn := 0; END_IF;
  910: (* FAULT: a step timed out, outputs off, alarm raised *)
      WdTime := T#0MS; Fault := TRUE; Busy := FALSE; Ready := FALSE;
      IF Ack AND Enable THEN Fault := FALSE; Sn := 10; END_IF;
END_CASE;
END_FUNCTION_BLOCK

(* oven door, Ofenschieber and lamp. Generated by stf-cad/hbw/sil/iec.py from the proven motion (control.py); do not edit. *)
FUNCTION_BLOCK FB_Door
VAR_INPUT
    Enable : BOOL;        (* K0 safety relay OK AND mode = AUTO *)
    Ack : BOOL;           (* HMI acknowledge *)
    Reset : BOOL;         (* S3 reset, via the safety relay *)
    Cmd : INT;            (* job to start (0 = none), taken when READY *)
    Arg1 : INT;           (* binding: slot / bay / slot pair index *)
    I6 : BOOL;           (* oven feeder inside *)
    I7 : BOOL;           (* oven feeder outside *)
    I10 : BOOL;           (* reed switch: oven door open *)
    I11 : BOOL;           (* reed switch: oven door shut *)
END_VAR
VAR_OUTPUT
    Q5 : BOOL;           (* oven feeder retract (M4) *)
    Q6 : BOOL;           (* oven feeder extend (M4) *)
    Q9 : BOOL;           (* oven lamp *)
    Q13 : BOOL;           (*  *)
    Ready, Busy, Done, Fault : BOOL;   (* Done: one scan, when a job ends *)
    Alarm : INT;          (* the state whose watchdog tripped *)
    Sn : INT;             (* the active state *)
END_VAR
VAR
    Prev : INT := -1;
    Job, B1 : INT;
    Wd : TON;             (* step watchdog *)
    Tm : TON;             (* step timer *)
    WdTime : TIME;        (* the active state's watchdog; 0 = none *)
END_VAR

(* every scan: outputs off unless the active state sets them; Done is a pulse *)
Q5 := FALSE; Q6 := FALSE; Q9 := FALSE; Q13 := FALSE; Done := FALSE;
IF NOT Enable AND Sn <> 900 THEN Sn := 900; END_IF;
Wd(IN := (Sn = Prev) AND (WdTime > T#0MS), PT := WdTime);
Tm(IN := (Sn = Prev), PT := T#1H);
Prev := Sn;
IF Wd.Q THEN Alarm := Sn; Sn := 910; END_IF;

CASE Sn OF
  0: (* INIT: power-up, all outputs off *)
      WdTime := T#0MS; IF Enable THEN Sn := 10; END_IF;
  10: (* H:open: door open *)
      WdTime := T#2000MS;
      Q13 := TRUE;
      IF I10 THEN Sn := 11; END_IF;
  11: (* H:slider: Ofenschieber in *)
      WdTime := T#3500MS;
      Q13 := TRUE; Q5 := TRUE;
      IF I6 THEN Sn := 12; END_IF;
  12: (* H:shut: door shut *)
      WdTime := T#2000MS;
      IF I11 THEN Sn := 100; END_IF;
  100: (* READY: homed, waiting for a job *)
      WdTime := T#0MS; Ready := TRUE; Busy := FALSE;
      IF Cmd <> 0 THEN Job := Cmd; B1 := Arg1; Busy := TRUE; Ready := FALSE;
          CASE Cmd OF 4: Sn := 1000; 5: Sn := 2000; 6: Sn := 3000; ELSE Sn := 910; Alarm := -Cmd; END_CASE;
      END_IF;
  1000: (* to_tt.01 row14: slider retracts *)
      WdTime := T#3500MS;
      Q13 := TRUE; Q5 := TRUE;
      IF I6 THEN Sn := 1001; END_IF;
  1001: (* to_tt.02 row15: door shuts *)
      WdTime := T#2000MS;
      IF I11 THEN Done := TRUE; Busy := FALSE; Sn := 100; END_IF;
  2000: (* bake.01 row3: Q5: slider retracts into the oven *)
      WdTime := T#3500MS;
      Q13 := TRUE; Q5 := TRUE;
      IF I6 THEN Sn := 2001; END_IF;
  2001: (* bake.02 row4: door shuts - bake (Q9 lamp) *)
      WdTime := T#2000MS;
      IF I11 THEN Sn := 2002; END_IF;
  2002: (* bake.03 row5: baking *)
      WdTime := T#0MS;
      Q9 := TRUE;
      IF Tm.ET >= T#2000MS THEN Sn := 2003; END_IF;
  2003: (* bake.04 row6: door opens *)
      WdTime := T#2000MS;
      Q13 := TRUE;
      IF I10 THEN Sn := 2004; END_IF;
  2004: (* bake.05 row7: slider extends *)
      WdTime := T#3500MS;
      Q13 := TRUE; Q6 := TRUE;
      IF I7 THEN Done := TRUE; Busy := FALSE; Sn := 100; END_IF;
  3000: (* present.01 row1: Q13: door opens *)
      WdTime := T#2000MS;
      Q13 := TRUE;
      IF I10 THEN Sn := 3001; END_IF;
  3001: (* present.02 row2: Q6: Ofenschieber extends - the VGR lays the workpiece on it (I9 breaks) *)
      WdTime := T#3500MS;
      Q13 := TRUE; Q6 := TRUE;
      IF I7 THEN Done := TRUE; Busy := FALSE; Sn := 100; END_IF;
  900: (* ESTOP: the safety relay dropped, outputs off *)
      WdTime := T#0MS; Busy := FALSE; Ready := FALSE; IF Reset AND Enable THEN Sn := 0; END_IF;
  910: (* FAULT: a step timed out, outputs off, alarm raised *)
      WdTime := T#0MS; Fault := TRUE; Busy := FALSE; Ready := FALSE;
      IF Ack AND Enable THEN Fault := FALSE; Sn := 10; END_IF;
END_CASE;
IF NOT I6 AND Sn <> 900 AND Sn <> 910 THEN Q13 := TRUE; END_IF;   (* F8: never shut on the Ofenschieber *)
END_FUNCTION_BLOCK

(* oven Sauggreifer. Generated by stf-cad/hbw/sil/iec.py from the proven motion (control.py); do not edit. *)
FUNCTION_BLOCK FB_Sauger
VAR_INPUT
    Enable : BOOL;        (* K0 safety relay OK AND mode = AUTO *)
    Ack : BOOL;           (* HMI acknowledge *)
    Reset : BOOL;         (* S3 reset, via the safety relay *)
    Cmd : INT;            (* job to start (0 = none), taken when READY *)
    Arg1 : INT;           (* binding: slot / bay / slot pair index *)
    I5 : BOOL;           (* reference vacuum (turntable position) *)
    I8 : BOOL;           (* vacuum at oven *)
    I12 : BOOL;           (* reed switch: Sauger lowered *)
    I13 : BOOL;           (* reed switch: Sauger up *)
END_VAR
VAR_OUTPUT
    Q7 : BOOL;           (* vacuum towards oven (M5) *)
    Q8 : BOOL;           (* vacuum towards turntable (M5) *)
    Q11 : BOOL;           (*  *)
    Q12 : BOOL;           (*  *)
    Ready, Busy, Done, Fault : BOOL;   (* Done: one scan, when a job ends *)
    Alarm : INT;          (* the state whose watchdog tripped *)
    Sn : INT;             (* the active state *)
END_VAR
VAR
    Prev : INT := -1;
    Job, B1 : INT;
    Wd : TON;             (* step watchdog *)
    Tm : TON;             (* step timer *)
    WdTime : TIME;        (* the active state's watchdog; 0 = none *)
END_VAR

(* every scan: outputs off unless the active state sets them; Done is a pulse *)
Q7 := FALSE; Q8 := FALSE; Q11 := FALSE; Q12 := FALSE; Done := FALSE;
IF NOT Enable AND Sn <> 900 THEN Sn := 900; END_IF;
Wd(IN := (Sn = Prev) AND (WdTime > T#0MS), PT := WdTime);
Tm(IN := (Sn = Prev), PT := T#1H);
Prev := Sn;
IF Wd.Q THEN Alarm := Sn; Sn := 910; END_IF;

CASE Sn OF
  0: (* INIT: power-up, all outputs off *)
      WdTime := T#0MS; IF Enable THEN Sn := 10; END_IF;
  10: (* H:up: Sauger up, vacuum off *)
      WdTime := T#1400MS;
      IF I13 THEN Sn := 11; END_IF;
  11: (* H:tt: Sauger to the Drehtisch *)
      WdTime := T#3500MS;
      Q8 := TRUE;
      IF I5 THEN Sn := 100; END_IF;
  100: (* READY: homed, waiting for a job *)
      WdTime := T#0MS; Ready := TRUE; Busy := FALSE;
      IF Cmd <> 0 THEN Job := Cmd; B1 := Arg1; Busy := TRUE; Ready := FALSE;
          CASE Cmd OF 4: Sn := 1000; ELSE Sn := 910; Alarm := -Cmd; END_CASE;
      END_IF;
  1000: (* to_tt.01 row8: Q7: Sauger to the oven (I8) *)
      WdTime := T#3500MS;
      Q7 := TRUE;
      IF I8 THEN Sn := 1001; END_IF;
  1001: (* to_tt.02 row9: Q12: lower onto the workpiece, Q11 vacuum *)
      WdTime := T#1400MS;
      Q11 := TRUE; Q12 := TRUE;
      IF I12 THEN Sn := 1002; END_IF;
  1002: (* to_tt.03 row10: lift *)
      WdTime := T#1400MS;
      Q11 := TRUE;
      IF I13 THEN Sn := 1003; END_IF;
  1003: (* to_tt.04 row11: Q8: Sauger to the Drehtisch (I5) *)
      WdTime := T#3500MS;
      Q11 := TRUE; Q8 := TRUE;
      IF I5 THEN Sn := 1004; END_IF;
  1004: (* to_tt.05 row12: lower, release onto the disc *)
      WdTime := T#1400MS;
      Q12 := TRUE;
      IF I12 THEN Sn := 1005; END_IF;
  1005: (* to_tt.06 row13: lift *)
      WdTime := T#1400MS;
      IF I13 THEN Done := TRUE; Busy := FALSE; Sn := 100; END_IF;
  900: (* ESTOP: the safety relay dropped, outputs off *)
      WdTime := T#0MS; Busy := FALSE; Ready := FALSE; IF Reset AND Enable THEN Sn := 0; END_IF;
  910: (* FAULT: a step timed out, outputs off, alarm raised *)
      WdTime := T#0MS; Fault := TRUE; Busy := FALSE; Ready := FALSE;
      IF Ack AND Enable THEN Fault := FALSE; Sn := 10; END_IF;
END_CASE;
END_FUNCTION_BLOCK

(* Drehtisch, Saege and Auswerfer. Generated by stf-cad/hbw/sil/iec.py from the proven motion (control.py); do not edit. *)
FUNCTION_BLOCK FB_Turntable
VAR_INPUT
    Enable : BOOL;        (* K0 safety relay OK AND mode = AUTO *)
    Ack : BOOL;           (* HMI acknowledge *)
    Reset : BOOL;         (* S3 reset, via the safety relay *)
    Cmd : INT;            (* job to start (0 = none), taken when READY *)
    Arg1 : INT;           (* binding: slot / bay / slot pair index *)
    I1 : BOOL;           (* reference turntable (vacuum position) *)
    I2 : BOOL;           (* reference turntable (belt position) *)
    I4 : BOOL;           (* reference turntable (saw position) *)
    I14 : BOOL;           (* reed switch: Auswerfer out *)
    I15 : BOOL;           (* reed switch: Auswerfer home *)
END_VAR
VAR_OUTPUT
    Q1 : BOOL;           (* turntable clockwise (M1) *)
    Q2 : BOOL;           (* turntable counter-clockwise (M1) *)
    Q4 : BOOL;           (* saw (M3) *)
    Q14 : BOOL;           (*  *)
    Ready, Busy, Done, Fault : BOOL;   (* Done: one scan, when a job ends *)
    Alarm : INT;          (* the state whose watchdog tripped *)
    Sn : INT;             (* the active state *)
END_VAR
VAR
    Prev : INT := -1;
    Job, B1 : INT;
    Wd : TON;             (* step watchdog *)
    Tm : TON;             (* step timer *)
    WdTime : TIME;        (* the active state's watchdog; 0 = none *)
END_VAR

(* every scan: outputs off unless the active state sets them; Done is a pulse *)
Q1 := FALSE; Q2 := FALSE; Q4 := FALSE; Q14 := FALSE; Done := FALSE;
IF NOT Enable AND Sn <> 900 THEN Sn := 900; END_IF;
Wd(IN := (Sn = Prev) AND (WdTime > T#0MS), PT := WdTime);
Tm(IN := (Sn = Prev), PT := T#1H);
Prev := Sn;
IF Wd.Q THEN Alarm := Sn; Sn := 910; END_IF;

CASE Sn OF
  0: (* INIT: power-up, all outputs off *)
      WdTime := T#0MS; IF Enable THEN Sn := 10; END_IF;
  10: (* H:push: Auswerfer home *)
      WdTime := T#1400MS;
      IF I15 THEN Sn := 11; END_IF;
  11: (* H:turn: Drehtisch to the vacuum position *)
      WdTime := T#2800MS;
      Q2 := TRUE;
      IF I1 THEN Sn := 100; END_IF;
  100: (* READY: homed, waiting for a job *)
      WdTime := T#0MS; Ready := TRUE; Busy := FALSE;
      IF Cmd <> 0 THEN Job := Cmd; B1 := Arg1; Busy := TRUE; Ready := FALSE;
          CASE Cmd OF 3: Sn := 1000; ELSE Sn := 910; Alarm := -Cmd; END_CASE;
      END_IF;
  1000: (* saw_eject.01 row16: Q1: Drehtisch to the Säge (I4) *)
      WdTime := T#2800MS;
      Q1 := TRUE;
      IF I4 THEN Sn := 1001; END_IF;
  1001: (* saw_eject.02 row17: Q4: saw runs *)
      WdTime := T#0MS;
      Q4 := TRUE;
      IF Tm.ET >= T#2000MS THEN Sn := 1002; END_IF;
  1002: (* saw_eject.03 row18: Drehtisch to the belt (I2) *)
      WdTime := T#2800MS;
      Q1 := TRUE;
      IF I2 THEN Sn := 1003; END_IF;
  1003: (* saw_eject.04 row19: Q14: Auswerfer pushes the workpiece onto the belt *)
      WdTime := T#1400MS;
      Q14 := TRUE;
      IF I14 THEN Sn := 1004; END_IF;
  1004: (* saw_eject.05 row20: Auswerfer home *)
      WdTime := T#1400MS;
      IF I15 THEN Sn := 1005; END_IF;
  1005: (* saw_eject.06 row21: I3 passed: Drehtisch home *)
      WdTime := T#5000MS;
      Q2 := TRUE;
      IF I1 THEN Done := TRUE; Busy := FALSE; Sn := 100; END_IF;
  900: (* ESTOP: the safety relay dropped, outputs off *)
      WdTime := T#0MS; Busy := FALSE; Ready := FALSE; IF Reset AND Enable THEN Sn := 0; END_IF;
  910: (* FAULT: a step timed out, outputs off, alarm raised *)
      WdTime := T#0MS; Fault := TRUE; Busy := FALSE; Ready := FALSE;
      IF Ack AND Enable THEN Fault := FALSE; Sn := 10; END_IF;
END_CASE;
END_FUNCTION_BLOCK

(* oven belt. Generated by stf-cad/hbw/sil/iec.py from the proven motion (control.py); do not edit. *)
FUNCTION_BLOCK FB_Ovenbelt
VAR_INPUT
    Enable : BOOL;        (* K0 safety relay OK AND mode = AUTO *)
    Ack : BOOL;           (* HMI acknowledge *)
    Reset : BOOL;         (* S3 reset, via the safety relay *)
    Cmd : INT;            (* job to start (0 = none), taken when READY *)
    Arg1 : INT;           (* binding: slot / bay / slot pair index *)
    I3 : BOOL;           (* light barrier end of conveyor belt *)
END_VAR
VAR_OUTPUT
    Q3 : BOOL;           (* conveyor belt (M2) *)
    Ready, Busy, Done, Fault : BOOL;   (* Done: one scan, when a job ends *)
    Alarm : INT;          (* the state whose watchdog tripped *)
    Sn : INT;             (* the active state *)
END_VAR
VAR
    Prev : INT := -1;
    Job, B1 : INT;
    Wd : TON;             (* step watchdog *)
    Tm : TON;             (* step timer *)
    WdTime : TIME;        (* the active state's watchdog; 0 = none *)
END_VAR

(* every scan: outputs off unless the active state sets them; Done is a pulse *)
Q3 := FALSE; Done := FALSE;
IF NOT Enable AND Sn <> 900 THEN Sn := 900; END_IF;
Wd(IN := (Sn = Prev) AND (WdTime > T#0MS), PT := WdTime);
Tm(IN := (Sn = Prev), PT := T#1H);
Prev := Sn;
IF Wd.Q THEN Alarm := Sn; Sn := 910; END_IF;

CASE Sn OF
  0: (* INIT: power-up, all outputs off *)
      WdTime := T#0MS; IF Enable THEN Sn := 100; END_IF;
  100: (* READY: homed, waiting for a job *)
      WdTime := T#0MS; Ready := TRUE; Busy := FALSE;
      IF Cmd <> 0 THEN Job := Cmd; B1 := Arg1; Busy := TRUE; Ready := FALSE;
          CASE Cmd OF 2: Sn := 1000; ELSE Sn := 910; Alarm := -Cmd; END_CASE;
      END_IF;
  1000: (* ovenbelt.01 run->I3: Q3 carries the cookie to I3 and onto the sorting inlet *)
      WdTime := T#9200MS;
      Q3 := TRUE;
      IF I3 THEN Done := TRUE; Busy := FALSE; Sn := 100; END_IF;
  900: (* ESTOP: the safety relay dropped, outputs off *)
      WdTime := T#0MS; Busy := FALSE; Ready := FALSE; IF Reset AND Enable THEN Sn := 0; END_IF;
  910: (* FAULT: a step timed out, outputs off, alarm raised *)
      WdTime := T#0MS; Fault := TRUE; Busy := FALSE; Ready := FALSE;
      IF Ack AND Enable THEN Fault := FALSE; Sn := 100; END_IF;
END_CASE;
END_FUNCTION_BLOCK

(* sorting line and ejectors. Generated by stf-cad/hbw/sil/iec.py from the proven motion (control.py); do not edit. *)
FUNCTION_BLOCK FB_Line
VAR_INPUT
    Enable : BOOL;        (* K0 safety relay OK AND mode = AUTO *)
    Ack : BOOL;           (* HMI acknowledge *)
    Reset : BOOL;         (* S3 reset, via the safety relay *)
    Cmd : INT;            (* job to start (0 = none), taken when READY *)
    Arg1 : INT;           (* binding: slot / bay / slot pair index *)
    I1 : BOOL;           (* pulse counter (Impulstaster) *)
    I3 : BOOL;           (* light barrier behind colour sensor *)
    I5 : BOOL;           (* light barrier white *)
    I6 : BOOL;           (* light barrier red *)
    I7 : BOOL;           (* light barrier blue *)
    A4 : INT;             (* colour sensor, mV *)
END_VAR
VAR_OUTPUT
    Q1 : BOOL;           (* conveyor belt *)
    Q3 : BOOL;           (*  *)
    Q4 : BOOL;           (*  *)
    Q5 : BOOL;           (*  *)
    Ready, Busy, Done, Fault : BOOL;   (* Done: one scan, when a job ends *)
    Alarm : INT;          (* the state whose watchdog tripped *)
    Sn : INT;             (* the active state *)
END_VAR
VAR
    Prev : INT := -1;
    Job, B1 : INT;
    Wd : TON;             (* step watchdog *)
    Tm : TON;             (* step timer *)
    WdTime : TIME;        (* the active state's watchdog; 0 = none *)
    MinMv : INT := 32767;
    Cls : INT;
    Pulses : INT;
    Edge : R_TRIG;
    Bar : BOOL;
END_VAR
VAR CONSTANT
    WD_SORT : ARRAY[1..3, 1..5] OF TIME := [T#6500MS, T#0MS, T#4100MS, T#1200MS, T#0MS, T#6500MS, T#0MS, T#8300MS, T#1200MS, T#0MS, T#6500MS, T#0MS, T#12500MS, T#1200MS, T#0MS];
    NEJECT : ARRAY[1..3] OF INT := [24, 52, 80];  (* I1 pulses from I3 to each ejector, 5 mm per pulse (ASSUMED) *)
END_VAR

(* every scan: outputs off unless the active state sets them; Done is a pulse *)
Q1 := FALSE; Q3 := FALSE; Q4 := FALSE; Q5 := FALSE; Done := FALSE;
IF NOT Enable AND Sn <> 900 THEN Sn := 900; END_IF;
Wd(IN := (Sn = Prev) AND (WdTime > T#0MS), PT := WdTime);
Tm(IN := (Sn = Prev), PT := T#1H);
Edge(CLK := I1);
IF Sn <> Prev THEN Pulses := 0; END_IF;
IF Edge.Q THEN Pulses := Pulses + 1; END_IF;
IF A4 < MinMv THEN MinMv := A4; END_IF;
CASE B1 OF 1: Bar := I5; 2: Bar := I6; 3: Bar := I7; ELSE Bar := FALSE; END_CASE;
Prev := Sn;
IF Wd.Q THEN Alarm := Sn; Sn := 910; END_IF;

CASE Sn OF
  0: (* INIT: power-up, all outputs off *)
      WdTime := T#0MS; IF Enable THEN Sn := 100; END_IF;
  100: (* READY: homed, waiting for a job *)
      WdTime := T#0MS; Ready := TRUE; Busy := FALSE;
      IF Cmd <> 0 THEN Job := Cmd; B1 := Arg1; Busy := TRUE; Ready := FALSE;
          CASE Cmd OF 1: Sn := 1000; ELSE Sn := 910; Alarm := -Cmd; END_CASE;
          MinMv := 32767;
      END_IF;
  1000: (* sort.01 run->I3: belt runs the cookie past the colour sensor; A4 sampled until I3 *)
      WdTime := T#6500MS;
      Q1 := TRUE;
      IF I3 THEN Sn := 1001; END_IF;
  1001: (* sort.02 classify: min(A4) over the pass -> flavour class; compared with the record *)
      WdTime := T#0MS;
      Q1 := TRUE;
      IF MinMv < 645 THEN Cls := 3;  ELSIF MinMv < 1305 THEN Cls := 2;  ELSE Cls := 1; END_IF;
      IF Cls = B1 THEN Sn := 1002; END_IF;
  1002: (* sort.03 run->eject: belt runs on; I1 pulses counted to the ejector *)
      WdTime := WD_SORT[B1, 3];
      Q1 := TRUE;
      IF Pulses >= NEJECT[B1] THEN Sn := 1003; END_IF;
  1003: (* sort.04 eject: belt stops; the ejector pushes the cookie into its bay *)
      WdTime := T#1200MS;
      CASE B1 OF 1: Q3 := TRUE; 2: Q4 := TRUE; 3: Q5 := TRUE; END_CASE;
      IF Bar THEN Sn := 1004; END_IF;
  1004: (* sort.05 eject_back: ejector back *)
      WdTime := T#0MS;
      IF Tm.ET >= T#500MS THEN Done := TRUE; Busy := FALSE; Sn := 100; END_IF;
  900: (* ESTOP: the safety relay dropped, outputs off *)
      WdTime := T#0MS; Busy := FALSE; Ready := FALSE; IF Reset AND Enable THEN Sn := 0; END_IF;
  910: (* FAULT: a step timed out, outputs off, alarm raised *)
      WdTime := T#0MS; Fault := TRUE; Busy := FALSE; Ready := FALSE;
      IF Ack AND Enable THEN Fault := FALSE; Sn := 100; END_IF;
END_CASE;
END_FUNCTION_BLOCK

(* The orchestrator: control.py's dispatcher, statement for statement. Generated by sil/iec.py. *)
PROGRAM MAIN
VAR
    hbw_I1 AT %IX0.0 : BOOL;
    hbw_I4 AT %IX0.1 : BOOL;
    hbw_I5 AT %IX0.2 : BOOL;
    hbw_I6 AT %IX0.3 : BOOL;
    hbw_I2 AT %IX0.4 : BOOL;
    hbw_I3 AT %IX0.5 : BOOL;
    vgr_I1 AT %IX0.6 : BOOL;
    vgr_I2 AT %IX0.7 : BOOL;
    vgr_I3 AT %IX1.0 : BOOL;
    vgr_I4 AT %IX1.1 : BOOL;
    oven_I6 AT %IX1.2 : BOOL;
    oven_I7 AT %IX1.3 : BOOL;
    oven_I10 AT %IX1.4 : BOOL;
    oven_I11 AT %IX1.5 : BOOL;
    oven_I5 AT %IX1.6 : BOOL;
    oven_I8 AT %IX1.7 : BOOL;
    oven_I12 AT %IX2.0 : BOOL;
    oven_I13 AT %IX2.1 : BOOL;
    oven_I1 AT %IX2.2 : BOOL;
    oven_I2 AT %IX2.3 : BOOL;
    oven_I4 AT %IX2.4 : BOOL;
    oven_I14 AT %IX2.5 : BOOL;
    oven_I15 AT %IX2.6 : BOOL;
    oven_I3 AT %IX2.7 : BOOL;
    sorting_I1 AT %IX3.0 : BOOL;
    sorting_I3 AT %IX3.1 : BOOL;
    sorting_I5 AT %IX3.2 : BOOL;
    sorting_I6 AT %IX3.3 : BOOL;
    sorting_I7 AT %IX3.4 : BOOL;
    hbw_RF1_Valid AT %IX3.5 : BOOL;
    hbw_RF2_Valid AT %IX3.6 : BOOL;
    cell_SafetyOK AT %IX3.7 : BOOL;
    hbw_RF2_Tag AT %IW0 : INT;
    sorting_A4 AT %IW1 : INT;
    hbw_PosTravel AT %ID0 : REAL;
    hbw_PosLift AT %ID1 : REAL;
    vgr_PosPlunge AT %ID2 : REAL;
    vgr_PosReach AT %ID3 : REAL;
    vgr_PosSwivel AT %ID4 : REAL;
    hbw_Q3 AT %QX0.0 : BOOL;
    hbw_Q4 AT %QX0.1 : BOOL;
    hbw_Q5 AT %QX0.2 : BOOL;
    hbw_Q6 AT %QX0.3 : BOOL;
    hbw_Q7 AT %QX0.4 : BOOL;
    hbw_Q8 AT %QX0.5 : BOOL;
    hbw_Q1 AT %QX0.6 : BOOL;
    hbw_Q2 AT %QX0.7 : BOOL;
    vgr_Q1 AT %QX1.0 : BOOL;
    vgr_Q2 AT %QX1.1 : BOOL;
    vgr_Q3 AT %QX1.2 : BOOL;
    vgr_Q4 AT %QX1.3 : BOOL;
    vgr_Q5 AT %QX1.4 : BOOL;
    vgr_Q6 AT %QX1.5 : BOOL;
    vgr_Q8 AT %QX1.6 : BOOL;
    oven_Q5 AT %QX1.7 : BOOL;
    oven_Q6 AT %QX2.0 : BOOL;
    oven_Q9 AT %QX2.1 : BOOL;
    oven_Q13 AT %QX2.2 : BOOL;
    oven_Q7 AT %QX2.3 : BOOL;
    oven_Q8 AT %QX2.4 : BOOL;
    oven_Q11 AT %QX2.5 : BOOL;
    oven_Q12 AT %QX2.6 : BOOL;
    oven_Q1 AT %QX2.7 : BOOL;
    oven_Q2 AT %QX3.0 : BOOL;
    oven_Q4 AT %QX3.1 : BOOL;
    oven_Q14 AT %QX3.2 : BOOL;
    oven_Q3 AT %QX3.3 : BOOL;
    sorting_Q1 AT %QX3.4 : BOOL;
    sorting_Q3 AT %QX3.5 : BOOL;
    sorting_Q4 AT %QX3.6 : BOOL;
    sorting_Q5 AT %QX3.7 : BOOL;
    mon_phase AT %MW0 : INT;
    mon_jobs AT %MW1 : INT;
    mon_crane_sn AT %MW10 : INT;
    mon_crane_job AT %MW11 : INT;
    mon_crane_b1 AT %MW12 : INT;
    mon_crane_b2 AT %MW13 : INT;
    mon_crane_b3 AT %MW14 : INT;
    mon_crane_b4 AT %MW15 : INT;
    mon_crane_b5 AT %MW16 : INT;
    mon_crane_b6 AT %MW17 : INT;
    mon_crane_alarm AT %MW18 : INT;
    mon_crane_seg AT %MW19 : INT;
    mon_crane_n AT %MW101 : INT;
    mon_belt_sn AT %MW20 : INT;
    mon_belt_job AT %MW21 : INT;
    mon_belt_b1 AT %MW22 : INT;
    mon_belt_b2 AT %MW23 : INT;
    mon_belt_b3 AT %MW24 : INT;
    mon_belt_b4 AT %MW25 : INT;
    mon_belt_b5 AT %MW26 : INT;
    mon_belt_b6 AT %MW27 : INT;
    mon_belt_alarm AT %MW28 : INT;
    mon_belt_seg AT %MW29 : INT;
    mon_belt_n AT %MW102 : INT;
    mon_arm_sn AT %MW30 : INT;
    mon_arm_job AT %MW31 : INT;
    mon_arm_b1 AT %MW32 : INT;
    mon_arm_b2 AT %MW33 : INT;
    mon_arm_b3 AT %MW34 : INT;
    mon_arm_b4 AT %MW35 : INT;
    mon_arm_b5 AT %MW36 : INT;
    mon_arm_b6 AT %MW37 : INT;
    mon_arm_alarm AT %MW38 : INT;
    mon_arm_seg AT %MW39 : INT;
    mon_arm_n AT %MW103 : INT;
    mon_door_sn AT %MW40 : INT;
    mon_door_job AT %MW41 : INT;
    mon_door_b1 AT %MW42 : INT;
    mon_door_b2 AT %MW43 : INT;
    mon_door_b3 AT %MW44 : INT;
    mon_door_b4 AT %MW45 : INT;
    mon_door_b5 AT %MW46 : INT;
    mon_door_b6 AT %MW47 : INT;
    mon_door_alarm AT %MW48 : INT;
    mon_door_seg AT %MW49 : INT;
    mon_door_n AT %MW104 : INT;
    mon_sauger_sn AT %MW50 : INT;
    mon_sauger_job AT %MW51 : INT;
    mon_sauger_b1 AT %MW52 : INT;
    mon_sauger_b2 AT %MW53 : INT;
    mon_sauger_b3 AT %MW54 : INT;
    mon_sauger_b4 AT %MW55 : INT;
    mon_sauger_b5 AT %MW56 : INT;
    mon_sauger_b6 AT %MW57 : INT;
    mon_sauger_alarm AT %MW58 : INT;
    mon_sauger_seg AT %MW59 : INT;
    mon_sauger_n AT %MW105 : INT;
    mon_turntable_sn AT %MW60 : INT;
    mon_turntable_job AT %MW61 : INT;
    mon_turntable_b1 AT %MW62 : INT;
    mon_turntable_b2 AT %MW63 : INT;
    mon_turntable_b3 AT %MW64 : INT;
    mon_turntable_b4 AT %MW65 : INT;
    mon_turntable_b5 AT %MW66 : INT;
    mon_turntable_b6 AT %MW67 : INT;
    mon_turntable_alarm AT %MW68 : INT;
    mon_turntable_seg AT %MW69 : INT;
    mon_turntable_n AT %MW106 : INT;
    mon_ovenbelt_sn AT %MW70 : INT;
    mon_ovenbelt_job AT %MW71 : INT;
    mon_ovenbelt_b1 AT %MW72 : INT;
    mon_ovenbelt_b2 AT %MW73 : INT;
    mon_ovenbelt_b3 AT %MW74 : INT;
    mon_ovenbelt_b4 AT %MW75 : INT;
    mon_ovenbelt_b5 AT %MW76 : INT;
    mon_ovenbelt_b6 AT %MW77 : INT;
    mon_ovenbelt_alarm AT %MW78 : INT;
    mon_ovenbelt_seg AT %MW79 : INT;
    mon_ovenbelt_n AT %MW107 : INT;
    mon_line_sn AT %MW80 : INT;
    mon_line_job AT %MW81 : INT;
    mon_line_b1 AT %MW82 : INT;
    mon_line_b2 AT %MW83 : INT;
    mon_line_b3 AT %MW84 : INT;
    mon_line_b4 AT %MW85 : INT;
    mon_line_b5 AT %MW86 : INT;
    mon_line_b6 AT %MW87 : INT;
    mon_line_alarm AT %MW88 : INT;
    mon_line_seg AT %MW89 : INT;
    mon_line_n AT %MW108 : INT;
END_VAR
VAR
    Crane : FB_Crane;
    Belt : FB_Belt;
    Arm : FB_Arm;
    Door : FB_Door;
    Sauger : FB_Sauger;
    Turntable : FB_Turntable;
    Ovenbelt : FB_Ovenbelt;
    Line : FB_Line;
    Cmd, Arg, RJ, Seg, Nst : ARRAY[1..8] OF INT;   (* per unit: command; per lead: job, segment, starts *)
    RB : ARRAY[1..8, 1..6] OF INT;                  (* per lead: the job's binding *)
    UBusy, Dn, Rdy : ARRAY[1..8] OF BOOL;
    BeltTag : INT;
    Phase, Jobs : INT;
    (* the factory, as control.py keeps it *)
    SlotM : ARRAY[1..12] OF INT := [1, 2, 3, 4, 5, 6, 7, 8, 9, 10, 11, 12];   (* mould in each slot, 0 = free *)
    SlotC : ARRAY[1..12] OF INT := [1, 2, 3, 4, 5, 6, 7, 8, 9, 0, 0, 0];   (* cookie in that mould *)
    BinM, BinC, BinMode, BoutM, BoutC, BoutMode : INT;   (* belt ends: mould, cookie, 1 out 2 fill 3 in *)
    Tray, Tt, Ovb, Inlet, CupC, CupSrc : INT;
    Tout : BOOL;
    Bay : ARRAY[1..3, 1..4] OF INT := [10, 0, 0, 0, 11, 0, 0, 0, 12, 0, 0, 0];
    BayN : ARRAY[1..3] OF INT := [1, 1, 1];
    Stage : ARRAY[1..12] OF INT := [1, 1, 1, 1, 1, 1, 1, 1, 1, 2, 2, 2];   (* 1 raw 2 return 3 returning 4 stored 5 baked 6 done *)
    (* reservations (destinations) and departures (sources) *)
    ResSlot, LvSlot : ARRAY[1..12] OF BOOL;
    ResBay : ARRAY[1..3] OF INT;
    LvBay : ARRAY[1..3] OF BOOL;
    ResBin, LvBin, ResBout, LvBout, ResTray, LvTray, ResTt, LvTt, ResOvb, LvOvb, ResSin, LvSin : BOOL;
    Started, Found : BOOL;
    i, j, k, n, c, b, m, tm, ts, Pend, jb : INT;
    x1, x2, x3, x4, x5, x6 : INT;
    BestT : REAL;
END_VAR
VAR CONSTANT
    FLV : ARRAY[1..12] OF INT := [3, 1, 2, 3, 1, 2, 3, 1, 2, 1, 2, 3];   (* cookie -> the bay of its flavour *)
    PROD : ARRAY[1..9] OF INT := [1, 2, 3, 4, 5, 6, 7, 8, 9];   (* production order *)
    ISRET : ARRAY[1..12] OF BOOL := [FALSE, FALSE, FALSE, FALSE, FALSE, FALSE, FALSE, FALSE, FALSE, TRUE, TRUE, TRUE];   (* a cookie that goes into the rack *)
    DUALT : ARRAY[1..12, 1..12] OF REAL := [0.0, 23.533, 23.533, 23.533, 22.383, 22.333, 22.333, 22.333, 22.783, 22.733, 22.733, 22.733, 23.533, 0.0, 21.933, 21.933, 22.333, 20.783, 20.733, 20.733, 22.733, 21.183, 21.133, 21.133, 23.533, 21.933, 0.0, 20.333, 22.333, 20.733, 19.183, 19.133, 22.733, 21.133, 19.583, 19.533, 23.533, 21.933, 20.333, 0.0, 22.333, 20.733, 19.133, 17.583, 22.733, 21.133, 19.533, 17.983, 22.383, 22.333, 22.333, 22.333, 0.0, 21.133, 21.133, 21.133, 21.583, 21.533, 21.533, 21.533, 22.333, 20.783, 20.733, 20.733, 21.133, 0.0, 19.533, 19.533, 21.533, 19.983, 19.933, 19.933, 22.333, 20.733, 19.183, 19.133, 21.133, 19.533, 0.0, 17.933, 21.533, 19.933, 18.383, 18.333, 22.333, 20.733, 19.133, 17.583, 21.133, 19.533, 17.933, 0.0, 21.533, 19.933, 18.333, 16.783, 22.783, 22.733, 22.733, 22.733, 21.583, 21.533, 21.533, 21.533, 0.0, 21.933, 21.933, 21.933, 22.733, 21.183, 21.133, 21.133, 21.533, 19.983, 19.933, 19.933, 21.933, 0.0, 20.333, 20.333, 22.733, 21.133, 19.583, 19.533, 21.533, 19.933, 18.383, 18.333, 21.933, 20.333, 0.0, 18.733, 22.733, 21.133, 19.533, 17.983, 21.533, 19.933, 18.333, 16.783, 21.933, 20.333, 18.733, 0.0];   (* dual-command trip, s *)
    BAYCAP : INT := 4;
END_VAR

(* 1. the unit sequencers, then their outputs *)
Crane(Enable := cell_SafetyOK, Ack := FALSE, Reset := FALSE, Cmd := Cmd[1], Arg1 := Arg[1], I1 := hbw_I1, I4 := hbw_I4, I5 := hbw_I5, I6 := hbw_I6, PosTravel := hbw_PosTravel, PosLift := hbw_PosLift);
IF Crane.Busy THEN Cmd[1] := 0; END_IF;
Dn[1] := Crane.Done; Rdy[1] := Crane.Ready;
hbw_Q3 := Crane.Q3; hbw_Q4 := Crane.Q4; hbw_Q5 := Crane.Q5; hbw_Q6 := Crane.Q6; hbw_Q7 := Crane.Q7; hbw_Q8 := Crane.Q8;
Belt(Enable := cell_SafetyOK, Ack := FALSE, Reset := FALSE, Cmd := Cmd[2], Arg1 := Arg[2], I2 := hbw_I2, I3 := hbw_I3, Tag := BeltTag, ExpI2 := FALSE, ExpI3 := FALSE, RF1_Valid := hbw_RF1_Valid, RF2_Valid := hbw_RF2_Valid, RF2_Tag := hbw_RF2_Tag);
IF Belt.Busy THEN Cmd[2] := 0; END_IF;
Dn[2] := Belt.Done; Rdy[2] := Belt.Ready;
hbw_Q1 := Belt.Q1; hbw_Q2 := Belt.Q2;
Arm(Enable := cell_SafetyOK, Ack := FALSE, Reset := FALSE, Cmd := Cmd[3], Arg1 := Arg[3], I1 := vgr_I1, I2 := vgr_I2, I3 := vgr_I3, I4 := vgr_I4, PosPlunge := vgr_PosPlunge, PosReach := vgr_PosReach, PosSwivel := vgr_PosSwivel);
IF Arm.Busy THEN Cmd[3] := 0; END_IF;
Dn[3] := Arm.Done; Rdy[3] := Arm.Ready;
vgr_Q1 := Arm.Q1; vgr_Q2 := Arm.Q2; vgr_Q3 := Arm.Q3; vgr_Q4 := Arm.Q4; vgr_Q5 := Arm.Q5; vgr_Q6 := Arm.Q6; vgr_Q8 := Arm.Q8;
Door(Enable := cell_SafetyOK, Ack := FALSE, Reset := FALSE, Cmd := Cmd[4], Arg1 := Arg[4], I6 := oven_I6, I7 := oven_I7, I10 := oven_I10, I11 := oven_I11);
IF Door.Busy THEN Cmd[4] := 0; END_IF;
Dn[4] := Door.Done; Rdy[4] := Door.Ready;
oven_Q5 := Door.Q5; oven_Q6 := Door.Q6; oven_Q9 := Door.Q9; oven_Q13 := Door.Q13;
Sauger(Enable := cell_SafetyOK, Ack := FALSE, Reset := FALSE, Cmd := Cmd[5], Arg1 := Arg[5], I5 := oven_I5, I8 := oven_I8, I12 := oven_I12, I13 := oven_I13);
IF Sauger.Busy THEN Cmd[5] := 0; END_IF;
Dn[5] := Sauger.Done; Rdy[5] := Sauger.Ready;
oven_Q7 := Sauger.Q7; oven_Q8 := Sauger.Q8; oven_Q11 := Sauger.Q11; oven_Q12 := Sauger.Q12;
Turntable(Enable := cell_SafetyOK, Ack := FALSE, Reset := FALSE, Cmd := Cmd[6], Arg1 := Arg[6], I1 := oven_I1, I2 := oven_I2, I4 := oven_I4, I14 := oven_I14, I15 := oven_I15);
IF Turntable.Busy THEN Cmd[6] := 0; END_IF;
Dn[6] := Turntable.Done; Rdy[6] := Turntable.Ready;
oven_Q1 := Turntable.Q1; oven_Q2 := Turntable.Q2; oven_Q4 := Turntable.Q4; oven_Q14 := Turntable.Q14;
Ovenbelt(Enable := cell_SafetyOK, Ack := FALSE, Reset := FALSE, Cmd := Cmd[7], Arg1 := Arg[7], I3 := oven_I3);
IF Ovenbelt.Busy THEN Cmd[7] := 0; END_IF;
Dn[7] := Ovenbelt.Done; Rdy[7] := Ovenbelt.Ready;
oven_Q3 := Ovenbelt.Q3;
Line(Enable := cell_SafetyOK, Ack := FALSE, Reset := FALSE, Cmd := Cmd[8], Arg1 := Arg[8], I1 := sorting_I1, I3 := sorting_I3, I5 := sorting_I5, I6 := sorting_I6, I7 := sorting_I7, A4 := sorting_A4);
IF Line.Busy THEN Cmd[8] := 0; END_IF;
Dn[8] := Line.Done; Rdy[8] := Line.Ready;
sorting_Q1 := Line.Q1; sorting_Q3 := Line.Q3; sorting_Q4 := Line.Q4; sorting_Q5 := Line.Q5;

(* 2. production starts once every unit has homed *)
IF Phase = 0 THEN
    Found := TRUE;
    FOR k := 1 TO 8 DO Found := Found AND Rdy[k]; END_FOR;
    IF Found THEN
        Phase := 1;
        REPEAT
            Started := FALSE;
            (* 1 sort: the cookie at the sorting inlet, if its bay has room *)
            IF NOT Started AND Inlet <> 0 AND NOT LvSin THEN
                b := FLV[Inlet];
                IF BayN[b] + ResBay[b] < BAYCAP AND NOT UBusy[8] THEN
                    (* start sort *)
                    UBusy[8] := TRUE;
                    RJ[8] := 1; Seg[8] := 8; Nst[8] := Nst[8] + 1;
                    RB[8, 1] := Inlet; RB[8, 2] := b; RB[8, 3] := 0; RB[8, 4] := 0; RB[8, 5] := 0; RB[8, 6] := 0;
                    Cmd[8] := 1; Arg[8] := b;
                    LvSin := TRUE; ResBay[b] := ResBay[b] + 1;
                    Started := TRUE;
                END_IF;
            END_IF;
            (* 2 oven belt -> sorting inlet *)
            IF NOT Started AND Ovb <> 0 AND NOT LvOvb AND NOT ResSin AND Inlet = 0 AND NOT UBusy[7] THEN
                (* start ovenbelt *)
                UBusy[7] := TRUE;
                RJ[7] := 2; Seg[7] := 7; Nst[7] := Nst[7] + 1;
                RB[7, 1] := Ovb; RB[7, 2] := 0; RB[7, 3] := 0; RB[7, 4] := 0; RB[7, 5] := 0; RB[7, 6] := 0;
                Cmd[7] := 2; Arg[7] := 1;
                LvOvb := TRUE; ResSin := TRUE;
                Started := TRUE;
            END_IF;
            (* 3 saw and eject *)
            IF NOT Started AND Tt <> 0 AND NOT LvTt AND Stage[Tt] = 5 AND NOT ResOvb AND Ovb = 0 AND NOT UBusy[6] THEN
                (* start saw_eject *)
                UBusy[6] := TRUE;
                RJ[6] := 3; Seg[6] := 6; Nst[6] := Nst[6] + 1;
                RB[6, 1] := Tt; RB[6, 2] := 0; RB[6, 3] := 0; RB[6, 4] := 0; RB[6, 5] := 0; RB[6, 6] := 0;
                Cmd[6] := 3; Arg[6] := 1;
                LvTt := TRUE; ResOvb := TRUE;
                Started := TRUE;
            END_IF;
            (* 4 Sauger: tray -> turntable *)
            IF NOT Started AND Tray <> 0 AND NOT LvTray AND Stage[Tray] = 5 AND NOT ResTt AND Tt = 0 AND NOT UBusy[5] AND NOT UBusy[4] THEN
                (* start to_tt *)
                UBusy[5] := TRUE; UBusy[4] := TRUE;
                RJ[5] := 4; Seg[5] := 5; Nst[5] := Nst[5] + 1;
                RB[5, 1] := Tray; RB[5, 2] := 0; RB[5, 3] := 0; RB[5, 4] := 0; RB[5, 5] := 0; RB[5, 6] := 0;
                Cmd[5] := 4; Arg[5] := 1;
                LvTray := TRUE; ResTt := TRUE;
                Started := TRUE;
            END_IF;
            (* 5 bake *)
            IF NOT Started AND Tray <> 0 AND NOT LvTray AND Stage[Tray] = 1 AND NOT UBusy[4] THEN
                (* start bake *)
                UBusy[4] := TRUE;
                RJ[4] := 5; Seg[4] := 4; Nst[4] := Nst[4] + 1;
                RB[4, 1] := Tray; RB[4, 2] := 0; RB[4, 3] := 0; RB[4, 4] := 0; RB[4, 5] := 0; RB[4, 6] := 0;
                Cmd[4] := 5; Arg[4] := 1;
                LvTray := TRUE;
                Started := TRUE;
            END_IF;
            (* 5a the oven presents its tray while the cookie for it is on its way *)
            IF NOT Started AND Tray = 0 AND NOT Tout AND (CupC <> 0 OR ResTray) AND NOT LvTray AND NOT UBusy[4] THEN
                (* start present *)
                UBusy[4] := TRUE;
                RJ[4] := 6; Seg[4] := 4; Nst[4] := Nst[4] + 1;
                RB[4, 1] := CupC; RB[4, 2] := 0; RB[4, 3] := 0; RB[4, 4] := 0; RB[4, 5] := 0; RB[4, 6] := 0;
                Cmd[4] := 6; Arg[4] := 1;
                Started := TRUE;
            END_IF;
            (* 5b the VGR lays the cookie on the presented tray *)
            IF NOT Started AND CupC <> 0 AND Tout AND Tray = 0 AND NOT UBusy[3] AND NOT UBusy[4] THEN
                (* start place_oven *)
                UBusy[3] := TRUE; UBusy[4] := TRUE;
                RJ[3] := 7; Seg[3] := 3; Nst[3] := Nst[3] + 1;
                RB[3, 1] := CupC; RB[3, 2] := CupSrc; RB[3, 3] := 0; RB[3, 4] := 0; RB[3, 5] := 0; RB[3, 6] := 0;
                Cmd[3] := 7; Arg[3] := 1;
                Started := TRUE;
            END_IF;
            (* 7 belt -> oven (the pick half): the oven is free of a committed cookie, the cup is empty *)
            IF NOT Started AND BoutM <> 0 AND BoutC <> 0 AND BoutMode = 1 AND NOT LvBout AND CupC = 0 AND NOT ResTray AND NOT UBusy[3] AND NOT UBusy[2] THEN
                (* start belt_to_oven *)
                UBusy[3] := TRUE; UBusy[2] := TRUE;
                RJ[3] := 8; Seg[3] := 3; Nst[3] := Nst[3] + 1;
                RB[3, 1] := BoutC; RB[3, 2] := BoutM; RB[3, 3] := 0; RB[3, 4] := 0; RB[3, 5] := 0; RB[3, 6] := 0;
                Cmd[3] := 8; Arg[3] := 1;
                LvBout := TRUE; ResTray := TRUE;
                Started := TRUE;
            END_IF;
            (* 9 bay -> the empty mould at the hand-over (the first bay holding a cookie that goes in) *)
            IF NOT Started AND BoutM <> 0 AND BoutC = 0 AND BoutMode = 2 AND NOT LvBout AND CupC = 0 THEN
                Found := FALSE;
                FOR i := 1 TO 3 DO
                    IF NOT Found THEN
                        FOR j := 1 TO BayN[i] DO
                            IF NOT Found AND Stage[Bay[i, j]] = 2 THEN Found := TRUE; c := Bay[i, j]; b := i; END_IF;
                        END_FOR;
                    END_IF;
                END_FOR;
                IF Found AND NOT UBusy[3] AND NOT UBusy[2] THEN
                    (* start bay_to_belt *)
                    UBusy[3] := TRUE; UBusy[2] := TRUE;
                    RJ[3] := 9; Seg[3] := 3; Nst[3] := Nst[3] + 1;
                    RB[3, 1] := c; RB[3, 2] := b; RB[3, 3] := BoutM; RB[3, 4] := 0; RB[3, 5] := 0; RB[3, 6] := 0;
                    Cmd[3] := 9; Arg[3] := b;
                    LvBay[b] := TRUE;
                    Started := TRUE;
                END_IF;
            END_IF;
            (* 10 belt back *)
            IF NOT Started AND BoutM <> 0 AND BoutMode = 3 AND NOT LvBout AND NOT ResBin AND BinM = 0 AND NOT UBusy[2] THEN
                (* start belt_back *)
                UBusy[2] := TRUE;
                RJ[2] := 10; Seg[2] := 2; Nst[2] := Nst[2] + 1;
                RB[2, 1] := BoutM; RB[2, 2] := BoutC; RB[2, 3] := 0; RB[2, 4] := 0; RB[2, 5] := 0; RB[2, 6] := 0;
                Cmd[2] := 10; Arg[2] := 1;
                LvBout := TRUE; ResBin := TRUE; BeltTag := BoutM;
                Started := TRUE;
            END_IF;
            (* the next cookie of the production order that is still raw in the rack, and its slot *)
            tm := 0; ts := 0;
            FOR i := 1 TO 9 DO
                IF tm = 0 AND Stage[PROD[i]] = 1 THEN
                    FOR j := 1 TO 12 DO IF SlotM[j] <> 0 AND SlotC[j] = PROD[i] THEN tm := PROD[i]; ts := j; END_IF; END_FOR;
                END_IF;
            END_FOR;
            (* 10a dual command: store the mould coming in in the free slot nearest the next cookie, retrieve that cookie *)
            IF NOT Started AND BinM <> 0 AND BinMode = 3 AND NOT LvBin AND tm <> 0 AND NOT ResBout AND BoutM = 0 THEN
                n := 0; BestT := 1.0E9;
                FOR i := 1 TO 12 DO
                    IF NOT ResSlot[i] AND SlotM[i] = 0 THEN
                        IF DUALT[i, ts] < BestT THEN BestT := DUALT[i, ts]; n := i; END_IF;
                    END_IF;
                END_FOR;
                IF n <> 0 AND NOT LvSlot[ts] AND NOT UBusy[1] AND NOT UBusy[2] THEN
                    (* start store_retrieve *)
                    UBusy[1] := TRUE; UBusy[2] := TRUE;
                    RJ[1] := 11; Seg[1] := 1; Nst[1] := Nst[1] + 1;
                    RB[1, 1] := BinM; RB[1, 2] := BinC; RB[1, 3] := n; RB[1, 4] := tm; RB[1, 5] := SlotM[ts]; RB[1, 6] := ts;
                    Cmd[1] := 11; Arg[1] := (n - 1) * 12 + ts;
                    LvBin := TRUE; LvSlot[ts] := TRUE; ResSlot[n] := TRUE; ResBin := TRUE;
                    Started := TRUE;
                END_IF;
            END_IF;
            (* 11 belt forward *)
            IF NOT Started AND BinM <> 0 AND (BinMode = 1 OR BinMode = 2) AND NOT LvBin AND NOT ResBout AND BoutM = 0 AND NOT UBusy[2] THEN
                (* start belt_fwd *)
                UBusy[2] := TRUE;
                RJ[2] := 12; Seg[2] := 2; Nst[2] := Nst[2] + 1;
                RB[2, 1] := BinM; RB[2, 2] := BinC; RB[2, 3] := 0; RB[2, 4] := 0; RB[2, 5] := 0; RB[2, 6] := 0;
                Cmd[2] := 12; Arg[2] := 1;
                LvBin := TRUE; ResBout := TRUE; BeltTag := BinM;
                Started := TRUE;
            END_IF;
            (* 12 store in the first free slot *)
            IF NOT Started AND BinM <> 0 AND BinMode = 3 AND NOT LvBin THEN
                n := 0;
                FOR i := 12 TO 1 BY -1 DO IF NOT ResSlot[i] AND SlotM[i] = 0 THEN n := i; END_IF; END_FOR;
                IF n <> 0 AND NOT UBusy[1] AND NOT UBusy[2] THEN
                    (* start store *)
                    UBusy[1] := TRUE; UBusy[2] := TRUE;
                    RJ[1] := 13; Seg[1] := 1; Nst[1] := Nst[1] + 1;
                    RB[1, 1] := BinM; RB[1, 2] := BinC; RB[1, 3] := n; RB[1, 4] := 0; RB[1, 5] := 0; RB[1, 6] := 0;
                    Cmd[1] := 13; Arg[1] := n;
                    LvBin := TRUE; ResSlot[n] := TRUE;
                    Started := TRUE;
                END_IF;
            END_IF;
            (* 13 fetch an empty mould for a cookie going in (with reuse: only when nothing is left to retrieve) *)
            IF NOT Started AND NOT ResBin AND BinM = 0 AND NOT ResBout AND BoutM = 0 AND tm = 0 THEN
                Pend := 0;
                FOR i := 1 TO 12 DO IF ISRET[i] AND Stage[i] = 2 THEN Pend := Pend + 1; END_IF; END_FOR;
                IF BinM <> 0 AND BinMode = 2 THEN Pend := Pend - 1; END_IF;
                IF BoutM <> 0 AND BoutMode = 2 THEN Pend := Pend - 1; END_IF;
                IF RJ[1] = 14 THEN Pend := Pend - 1; END_IF;
                IF Pend > 0 THEN
                    n := 0;
                    FOR i := 12 TO 1 BY -1 DO IF SlotM[i] <> 0 AND SlotC[i] = 0 AND NOT LvSlot[i] THEN n := i; END_IF; END_FOR;
                    IF n <> 0 AND NOT UBusy[1] AND NOT UBusy[2] THEN
                        (* start fetch_empty *)
                        UBusy[1] := TRUE; UBusy[2] := TRUE;
                        RJ[1] := 14; Seg[1] := 1; Nst[1] := Nst[1] + 1;
                        RB[1, 1] := SlotM[n]; RB[1, 2] := n; RB[1, 3] := 0; RB[1, 4] := 0; RB[1, 5] := 0; RB[1, 6] := 0;
                        Cmd[1] := 14; Arg[1] := n;
                        LvSlot[n] := TRUE; ResBin := TRUE;
                        Started := TRUE;
                    END_IF;
                END_IF;
            END_IF;
            (* 14 retrieve the next cookie in production order *)
            IF NOT Started AND NOT ResBin AND BinM = 0 AND NOT ResBout AND BoutM = 0 AND tm <> 0 THEN
                IF NOT LvSlot[ts] AND NOT UBusy[1] AND NOT UBusy[2] THEN
                    (* start retrieve *)
                    UBusy[1] := TRUE; UBusy[2] := TRUE;
                    RJ[1] := 15; Seg[1] := 1; Nst[1] := Nst[1] + 1;
                    RB[1, 1] := tm; RB[1, 2] := SlotM[ts]; RB[1, 3] := ts; RB[1, 4] := 0; RB[1, 5] := 0; RB[1, 6] := 0;
                    Cmd[1] := 15; Arg[1] := ts;
                    LvSlot[ts] := TRUE; ResBin := TRUE;
                    Started := TRUE;
                END_IF;
            END_IF;
        UNTIL NOT Started
        END_REPEAT;
    END_IF;
END_IF;

(* 3. completions, leads in unit order (control.simulate's tie order); each is followed by a dispatch *)
IF Phase = 1 THEN
    FOR k := 1 TO 8 DO
        IF RJ[k] <> 0 AND Seg[k] <> 0 THEN
            IF Dn[Seg[k]] THEN
                IF RJ[k] = 4 AND Seg[k] = 5 THEN   (* to_tt: next segment *)
                    Seg[k] := 4; Cmd[4] := 4; Arg[4] := Arg[5]; Dn[5] := FALSE;
                END_IF;
            END_IF;
            IF Dn[Seg[k]] THEN
                (* complete the job lead k runs: control.complete() *)
                jb := RJ[k]; x1 := RB[k, 1]; x2 := RB[k, 2]; x3 := RB[k, 3]; x4 := RB[k, 4]; x5 := RB[k, 5]; x6 := RB[k, 6];
                RJ[k] := 0; Seg[k] := 0; Jobs := Jobs + 1;
                CASE jb OF
                  1: (* sort *)
                      UBusy[8] := FALSE;
                      LvSin := FALSE; ResBay[x2] := ResBay[x2] - 1;
                      BayN[x2] := BayN[x2] + 1; Bay[x2, BayN[x2]] := x1; Inlet := 0; Stage[x1] := 6;
                  2: (* ovenbelt *)
                      UBusy[7] := FALSE;
                      LvOvb := FALSE; ResSin := FALSE;
                      Inlet := Ovb; Ovb := 0;
                  3: (* saw_eject *)
                      UBusy[6] := FALSE;
                      LvTt := FALSE; ResOvb := FALSE;
                      Ovb := Tt; Tt := 0; Stage[x1] := 5;
                  4: (* to_tt *)
                      UBusy[5] := FALSE; UBusy[4] := FALSE;
                      LvTray := FALSE; ResTt := FALSE;
                      Tt := Tray; Tray := 0; Tout := FALSE;
                  5: (* bake *)
                      UBusy[4] := FALSE;
                      LvTray := FALSE;
                      Stage[x1] := 5;
                  6: (* present *)
                      UBusy[4] := FALSE;
                      Tout := TRUE;
                  7: (* place_oven *)
                      UBusy[3] := FALSE; UBusy[4] := FALSE;
                      Tray := CupC; CupC := 0; CupSrc := 0;
                  8: (* belt_to_oven *)
                      UBusy[3] := FALSE; UBusy[2] := FALSE;
                      LvBout := FALSE; ResTray := FALSE;
                      Pend := 0;
                      FOR i := 1 TO 12 DO IF ISRET[i] AND Stage[i] = 2 THEN Pend := Pend + 1; END_IF; END_FOR;
                      IF BinM <> 0 AND BinMode = 2 THEN Pend := Pend - 1; END_IF;
                      IF BoutM <> 0 AND BoutMode = 2 THEN Pend := Pend - 1; END_IF;
                      IF RJ[1] = 14 THEN Pend := Pend - 1; END_IF;
                      BoutC := 0; IF Pend > 0 THEN BoutMode := 2; ELSE BoutMode := 3; END_IF;
                      CupC := x1; CupSrc := 1;
                  9: (* bay_to_belt *)
                      UBusy[3] := FALSE; UBusy[2] := FALSE;
                      LvBay[x2] := FALSE;
                      n := 0;
                      FOR j := 1 TO BayN[x2] DO IF Bay[x2, j] <> x1 THEN n := n + 1; Bay[x2, n] := Bay[x2, j]; END_IF; END_FOR;
                      FOR j := n + 1 TO BAYCAP DO Bay[x2, j] := 0; END_FOR;
                      BayN[x2] := n; BoutM := x3; BoutC := x1; BoutMode := 3; Stage[x1] := 3;
                  10: (* belt_back *)
                      UBusy[2] := FALSE;
                      LvBout := FALSE; ResBin := FALSE;
                      BinM := BoutM; BinC := BoutC; BinMode := BoutMode; BoutM := 0; BoutC := 0; BoutMode := 0;
                  11: (* store_retrieve *)
                      UBusy[1] := FALSE; UBusy[2] := FALSE;
                      LvBin := FALSE; LvSlot[x6] := FALSE; ResSlot[x3] := FALSE; ResBin := FALSE;
                      SlotM[x3] := x1; SlotC[x3] := x2; SlotM[x6] := 0; SlotC[x6] := 0;
                      IF x2 <> 0 THEN Stage[x2] := 4; END_IF;
                      BinM := x5; BinC := x4; BinMode := 1;
                  12: (* belt_fwd *)
                      UBusy[2] := FALSE;
                      LvBin := FALSE; ResBout := FALSE;
                      BoutM := BinM; BoutC := BinC; BoutMode := BinMode; BinM := 0; BinC := 0; BinMode := 0;
                  13: (* store *)
                      UBusy[1] := FALSE; UBusy[2] := FALSE;
                      LvBin := FALSE; ResSlot[x3] := FALSE;
                      SlotM[x3] := x1; SlotC[x3] := x2; BinM := 0; BinC := 0; BinMode := 0;
                      IF x2 <> 0 THEN Stage[x2] := 4; END_IF;
                  14: (* fetch_empty *)
                      UBusy[1] := FALSE; UBusy[2] := FALSE;
                      LvSlot[x2] := FALSE; ResBin := FALSE;
                      SlotM[x2] := 0; SlotC[x2] := 0; BinM := x1; BinC := 0; BinMode := 2;
                  15: (* retrieve *)
                      UBusy[1] := FALSE; UBusy[2] := FALSE;
                      LvSlot[x3] := FALSE; ResBin := FALSE;
                      SlotM[x3] := 0; SlotC[x3] := 0; BinM := x2; BinC := x1; BinMode := 1;
                END_CASE;
                REPEAT
                    Started := FALSE;
                    (* 1 sort: the cookie at the sorting inlet, if its bay has room *)
                    IF NOT Started AND Inlet <> 0 AND NOT LvSin THEN
                        b := FLV[Inlet];
                        IF BayN[b] + ResBay[b] < BAYCAP AND NOT UBusy[8] THEN
                            (* start sort *)
                            UBusy[8] := TRUE;
                            RJ[8] := 1; Seg[8] := 8; Nst[8] := Nst[8] + 1;
                            RB[8, 1] := Inlet; RB[8, 2] := b; RB[8, 3] := 0; RB[8, 4] := 0; RB[8, 5] := 0; RB[8, 6] := 0;
                            Cmd[8] := 1; Arg[8] := b;
                            LvSin := TRUE; ResBay[b] := ResBay[b] + 1;
                            Started := TRUE;
                        END_IF;
                    END_IF;
                    (* 2 oven belt -> sorting inlet *)
                    IF NOT Started AND Ovb <> 0 AND NOT LvOvb AND NOT ResSin AND Inlet = 0 AND NOT UBusy[7] THEN
                        (* start ovenbelt *)
                        UBusy[7] := TRUE;
                        RJ[7] := 2; Seg[7] := 7; Nst[7] := Nst[7] + 1;
                        RB[7, 1] := Ovb; RB[7, 2] := 0; RB[7, 3] := 0; RB[7, 4] := 0; RB[7, 5] := 0; RB[7, 6] := 0;
                        Cmd[7] := 2; Arg[7] := 1;
                        LvOvb := TRUE; ResSin := TRUE;
                        Started := TRUE;
                    END_IF;
                    (* 3 saw and eject *)
                    IF NOT Started AND Tt <> 0 AND NOT LvTt AND Stage[Tt] = 5 AND NOT ResOvb AND Ovb = 0 AND NOT UBusy[6] THEN
                        (* start saw_eject *)
                        UBusy[6] := TRUE;
                        RJ[6] := 3; Seg[6] := 6; Nst[6] := Nst[6] + 1;
                        RB[6, 1] := Tt; RB[6, 2] := 0; RB[6, 3] := 0; RB[6, 4] := 0; RB[6, 5] := 0; RB[6, 6] := 0;
                        Cmd[6] := 3; Arg[6] := 1;
                        LvTt := TRUE; ResOvb := TRUE;
                        Started := TRUE;
                    END_IF;
                    (* 4 Sauger: tray -> turntable *)
                    IF NOT Started AND Tray <> 0 AND NOT LvTray AND Stage[Tray] = 5 AND NOT ResTt AND Tt = 0 AND NOT UBusy[5] AND NOT UBusy[4] THEN
                        (* start to_tt *)
                        UBusy[5] := TRUE; UBusy[4] := TRUE;
                        RJ[5] := 4; Seg[5] := 5; Nst[5] := Nst[5] + 1;
                        RB[5, 1] := Tray; RB[5, 2] := 0; RB[5, 3] := 0; RB[5, 4] := 0; RB[5, 5] := 0; RB[5, 6] := 0;
                        Cmd[5] := 4; Arg[5] := 1;
                        LvTray := TRUE; ResTt := TRUE;
                        Started := TRUE;
                    END_IF;
                    (* 5 bake *)
                    IF NOT Started AND Tray <> 0 AND NOT LvTray AND Stage[Tray] = 1 AND NOT UBusy[4] THEN
                        (* start bake *)
                        UBusy[4] := TRUE;
                        RJ[4] := 5; Seg[4] := 4; Nst[4] := Nst[4] + 1;
                        RB[4, 1] := Tray; RB[4, 2] := 0; RB[4, 3] := 0; RB[4, 4] := 0; RB[4, 5] := 0; RB[4, 6] := 0;
                        Cmd[4] := 5; Arg[4] := 1;
                        LvTray := TRUE;
                        Started := TRUE;
                    END_IF;
                    (* 5a the oven presents its tray while the cookie for it is on its way *)
                    IF NOT Started AND Tray = 0 AND NOT Tout AND (CupC <> 0 OR ResTray) AND NOT LvTray AND NOT UBusy[4] THEN
                        (* start present *)
                        UBusy[4] := TRUE;
                        RJ[4] := 6; Seg[4] := 4; Nst[4] := Nst[4] + 1;
                        RB[4, 1] := CupC; RB[4, 2] := 0; RB[4, 3] := 0; RB[4, 4] := 0; RB[4, 5] := 0; RB[4, 6] := 0;
                        Cmd[4] := 6; Arg[4] := 1;
                        Started := TRUE;
                    END_IF;
                    (* 5b the VGR lays the cookie on the presented tray *)
                    IF NOT Started AND CupC <> 0 AND Tout AND Tray = 0 AND NOT UBusy[3] AND NOT UBusy[4] THEN
                        (* start place_oven *)
                        UBusy[3] := TRUE; UBusy[4] := TRUE;
                        RJ[3] := 7; Seg[3] := 3; Nst[3] := Nst[3] + 1;
                        RB[3, 1] := CupC; RB[3, 2] := CupSrc; RB[3, 3] := 0; RB[3, 4] := 0; RB[3, 5] := 0; RB[3, 6] := 0;
                        Cmd[3] := 7; Arg[3] := 1;
                        Started := TRUE;
                    END_IF;
                    (* 7 belt -> oven (the pick half): the oven is free of a committed cookie, the cup is empty *)
                    IF NOT Started AND BoutM <> 0 AND BoutC <> 0 AND BoutMode = 1 AND NOT LvBout AND CupC = 0 AND NOT ResTray AND NOT UBusy[3] AND NOT UBusy[2] THEN
                        (* start belt_to_oven *)
                        UBusy[3] := TRUE; UBusy[2] := TRUE;
                        RJ[3] := 8; Seg[3] := 3; Nst[3] := Nst[3] + 1;
                        RB[3, 1] := BoutC; RB[3, 2] := BoutM; RB[3, 3] := 0; RB[3, 4] := 0; RB[3, 5] := 0; RB[3, 6] := 0;
                        Cmd[3] := 8; Arg[3] := 1;
                        LvBout := TRUE; ResTray := TRUE;
                        Started := TRUE;
                    END_IF;
                    (* 9 bay -> the empty mould at the hand-over (the first bay holding a cookie that goes in) *)
                    IF NOT Started AND BoutM <> 0 AND BoutC = 0 AND BoutMode = 2 AND NOT LvBout AND CupC = 0 THEN
                        Found := FALSE;
                        FOR i := 1 TO 3 DO
                            IF NOT Found THEN
                                FOR j := 1 TO BayN[i] DO
                                    IF NOT Found AND Stage[Bay[i, j]] = 2 THEN Found := TRUE; c := Bay[i, j]; b := i; END_IF;
                                END_FOR;
                            END_IF;
                        END_FOR;
                        IF Found AND NOT UBusy[3] AND NOT UBusy[2] THEN
                            (* start bay_to_belt *)
                            UBusy[3] := TRUE; UBusy[2] := TRUE;
                            RJ[3] := 9; Seg[3] := 3; Nst[3] := Nst[3] + 1;
                            RB[3, 1] := c; RB[3, 2] := b; RB[3, 3] := BoutM; RB[3, 4] := 0; RB[3, 5] := 0; RB[3, 6] := 0;
                            Cmd[3] := 9; Arg[3] := b;
                            LvBay[b] := TRUE;
                            Started := TRUE;
                        END_IF;
                    END_IF;
                    (* 10 belt back *)
                    IF NOT Started AND BoutM <> 0 AND BoutMode = 3 AND NOT LvBout AND NOT ResBin AND BinM = 0 AND NOT UBusy[2] THEN
                        (* start belt_back *)
                        UBusy[2] := TRUE;
                        RJ[2] := 10; Seg[2] := 2; Nst[2] := Nst[2] + 1;
                        RB[2, 1] := BoutM; RB[2, 2] := BoutC; RB[2, 3] := 0; RB[2, 4] := 0; RB[2, 5] := 0; RB[2, 6] := 0;
                        Cmd[2] := 10; Arg[2] := 1;
                        LvBout := TRUE; ResBin := TRUE; BeltTag := BoutM;
                        Started := TRUE;
                    END_IF;
                    (* the next cookie of the production order that is still raw in the rack, and its slot *)
                    tm := 0; ts := 0;
                    FOR i := 1 TO 9 DO
                        IF tm = 0 AND Stage[PROD[i]] = 1 THEN
                            FOR j := 1 TO 12 DO IF SlotM[j] <> 0 AND SlotC[j] = PROD[i] THEN tm := PROD[i]; ts := j; END_IF; END_FOR;
                        END_IF;
                    END_FOR;
                    (* 10a dual command: store the mould coming in in the free slot nearest the next cookie, retrieve that cookie *)
                    IF NOT Started AND BinM <> 0 AND BinMode = 3 AND NOT LvBin AND tm <> 0 AND NOT ResBout AND BoutM = 0 THEN
                        n := 0; BestT := 1.0E9;
                        FOR i := 1 TO 12 DO
                            IF NOT ResSlot[i] AND SlotM[i] = 0 THEN
                                IF DUALT[i, ts] < BestT THEN BestT := DUALT[i, ts]; n := i; END_IF;
                            END_IF;
                        END_FOR;
                        IF n <> 0 AND NOT LvSlot[ts] AND NOT UBusy[1] AND NOT UBusy[2] THEN
                            (* start store_retrieve *)
                            UBusy[1] := TRUE; UBusy[2] := TRUE;
                            RJ[1] := 11; Seg[1] := 1; Nst[1] := Nst[1] + 1;
                            RB[1, 1] := BinM; RB[1, 2] := BinC; RB[1, 3] := n; RB[1, 4] := tm; RB[1, 5] := SlotM[ts]; RB[1, 6] := ts;
                            Cmd[1] := 11; Arg[1] := (n - 1) * 12 + ts;
                            LvBin := TRUE; LvSlot[ts] := TRUE; ResSlot[n] := TRUE; ResBin := TRUE;
                            Started := TRUE;
                        END_IF;
                    END_IF;
                    (* 11 belt forward *)
                    IF NOT Started AND BinM <> 0 AND (BinMode = 1 OR BinMode = 2) AND NOT LvBin AND NOT ResBout AND BoutM = 0 AND NOT UBusy[2] THEN
                        (* start belt_fwd *)
                        UBusy[2] := TRUE;
                        RJ[2] := 12; Seg[2] := 2; Nst[2] := Nst[2] + 1;
                        RB[2, 1] := BinM; RB[2, 2] := BinC; RB[2, 3] := 0; RB[2, 4] := 0; RB[2, 5] := 0; RB[2, 6] := 0;
                        Cmd[2] := 12; Arg[2] := 1;
                        LvBin := TRUE; ResBout := TRUE; BeltTag := BinM;
                        Started := TRUE;
                    END_IF;
                    (* 12 store in the first free slot *)
                    IF NOT Started AND BinM <> 0 AND BinMode = 3 AND NOT LvBin THEN
                        n := 0;
                        FOR i := 12 TO 1 BY -1 DO IF NOT ResSlot[i] AND SlotM[i] = 0 THEN n := i; END_IF; END_FOR;
                        IF n <> 0 AND NOT UBusy[1] AND NOT UBusy[2] THEN
                            (* start store *)
                            UBusy[1] := TRUE; UBusy[2] := TRUE;
                            RJ[1] := 13; Seg[1] := 1; Nst[1] := Nst[1] + 1;
                            RB[1, 1] := BinM; RB[1, 2] := BinC; RB[1, 3] := n; RB[1, 4] := 0; RB[1, 5] := 0; RB[1, 6] := 0;
                            Cmd[1] := 13; Arg[1] := n;
                            LvBin := TRUE; ResSlot[n] := TRUE;
                            Started := TRUE;
                        END_IF;
                    END_IF;
                    (* 13 fetch an empty mould for a cookie going in (with reuse: only when nothing is left to retrieve) *)
                    IF NOT Started AND NOT ResBin AND BinM = 0 AND NOT ResBout AND BoutM = 0 AND tm = 0 THEN
                        Pend := 0;
                        FOR i := 1 TO 12 DO IF ISRET[i] AND Stage[i] = 2 THEN Pend := Pend + 1; END_IF; END_FOR;
                        IF BinM <> 0 AND BinMode = 2 THEN Pend := Pend - 1; END_IF;
                        IF BoutM <> 0 AND BoutMode = 2 THEN Pend := Pend - 1; END_IF;
                        IF RJ[1] = 14 THEN Pend := Pend - 1; END_IF;
                        IF Pend > 0 THEN
                            n := 0;
                            FOR i := 12 TO 1 BY -1 DO IF SlotM[i] <> 0 AND SlotC[i] = 0 AND NOT LvSlot[i] THEN n := i; END_IF; END_FOR;
                            IF n <> 0 AND NOT UBusy[1] AND NOT UBusy[2] THEN
                                (* start fetch_empty *)
                                UBusy[1] := TRUE; UBusy[2] := TRUE;
                                RJ[1] := 14; Seg[1] := 1; Nst[1] := Nst[1] + 1;
                                RB[1, 1] := SlotM[n]; RB[1, 2] := n; RB[1, 3] := 0; RB[1, 4] := 0; RB[1, 5] := 0; RB[1, 6] := 0;
                                Cmd[1] := 14; Arg[1] := n;
                                LvSlot[n] := TRUE; ResBin := TRUE;
                                Started := TRUE;
                            END_IF;
                        END_IF;
                    END_IF;
                    (* 14 retrieve the next cookie in production order *)
                    IF NOT Started AND NOT ResBin AND BinM = 0 AND NOT ResBout AND BoutM = 0 AND tm <> 0 THEN
                        IF NOT LvSlot[ts] AND NOT UBusy[1] AND NOT UBusy[2] THEN
                            (* start retrieve *)
                            UBusy[1] := TRUE; UBusy[2] := TRUE;
                            RJ[1] := 15; Seg[1] := 1; Nst[1] := Nst[1] + 1;
                            RB[1, 1] := tm; RB[1, 2] := SlotM[ts]; RB[1, 3] := ts; RB[1, 4] := 0; RB[1, 5] := 0; RB[1, 6] := 0;
                            Cmd[1] := 15; Arg[1] := ts;
                            LvSlot[ts] := TRUE; ResBin := TRUE;
                            Started := TRUE;
                        END_IF;
                    END_IF;
                UNTIL NOT Started
                END_REPEAT;
            END_IF;
        END_IF;
    END_FOR;
    (* the order is complete: nothing running, nothing in transit, every cookie done or stored *)
    Found := (BinM = 0) AND (BoutM = 0) AND (Tray = 0) AND (Tt = 0) AND (Ovb = 0) AND (Inlet = 0) AND (CupC = 0);
    FOR k := 1 TO 8 DO Found := Found AND (RJ[k] = 0); END_FOR;
    FOR k := 1 TO 9 DO Found := Found AND (Stage[PROD[k]] = 6); END_FOR;
    IF Found THEN Phase := 2; END_IF;
END_IF;

(* 4. the monitor *)
mon_phase := Phase; mon_jobs := Jobs;
mon_crane_sn := Crane.Sn; mon_crane_job := RJ[1]; mon_crane_alarm := Crane.Alarm; mon_crane_seg := Seg[1]; mon_crane_n := Nst[1];
mon_crane_b1 := RB[1, 1]; mon_crane_b2 := RB[1, 2]; mon_crane_b3 := RB[1, 3]; mon_crane_b4 := RB[1, 4]; mon_crane_b5 := RB[1, 5]; mon_crane_b6 := RB[1, 6];
mon_belt_sn := Belt.Sn; mon_belt_job := RJ[2]; mon_belt_alarm := Belt.Alarm; mon_belt_seg := Seg[2]; mon_belt_n := Nst[2];
mon_belt_b1 := RB[2, 1]; mon_belt_b2 := RB[2, 2]; mon_belt_b3 := RB[2, 3]; mon_belt_b4 := RB[2, 4]; mon_belt_b5 := RB[2, 5]; mon_belt_b6 := RB[2, 6];
mon_arm_sn := Arm.Sn; mon_arm_job := RJ[3]; mon_arm_alarm := Arm.Alarm; mon_arm_seg := Seg[3]; mon_arm_n := Nst[3];
mon_arm_b1 := RB[3, 1]; mon_arm_b2 := RB[3, 2]; mon_arm_b3 := RB[3, 3]; mon_arm_b4 := RB[3, 4]; mon_arm_b5 := RB[3, 5]; mon_arm_b6 := RB[3, 6];
mon_door_sn := Door.Sn; mon_door_job := RJ[4]; mon_door_alarm := Door.Alarm; mon_door_seg := Seg[4]; mon_door_n := Nst[4];
mon_door_b1 := RB[4, 1]; mon_door_b2 := RB[4, 2]; mon_door_b3 := RB[4, 3]; mon_door_b4 := RB[4, 4]; mon_door_b5 := RB[4, 5]; mon_door_b6 := RB[4, 6];
mon_sauger_sn := Sauger.Sn; mon_sauger_job := RJ[5]; mon_sauger_alarm := Sauger.Alarm; mon_sauger_seg := Seg[5]; mon_sauger_n := Nst[5];
mon_sauger_b1 := RB[5, 1]; mon_sauger_b2 := RB[5, 2]; mon_sauger_b3 := RB[5, 3]; mon_sauger_b4 := RB[5, 4]; mon_sauger_b5 := RB[5, 5]; mon_sauger_b6 := RB[5, 6];
mon_turntable_sn := Turntable.Sn; mon_turntable_job := RJ[6]; mon_turntable_alarm := Turntable.Alarm; mon_turntable_seg := Seg[6]; mon_turntable_n := Nst[6];
mon_turntable_b1 := RB[6, 1]; mon_turntable_b2 := RB[6, 2]; mon_turntable_b3 := RB[6, 3]; mon_turntable_b4 := RB[6, 4]; mon_turntable_b5 := RB[6, 5]; mon_turntable_b6 := RB[6, 6];
mon_ovenbelt_sn := Ovenbelt.Sn; mon_ovenbelt_job := RJ[7]; mon_ovenbelt_alarm := Ovenbelt.Alarm; mon_ovenbelt_seg := Seg[7]; mon_ovenbelt_n := Nst[7];
mon_ovenbelt_b1 := RB[7, 1]; mon_ovenbelt_b2 := RB[7, 2]; mon_ovenbelt_b3 := RB[7, 3]; mon_ovenbelt_b4 := RB[7, 4]; mon_ovenbelt_b5 := RB[7, 5]; mon_ovenbelt_b6 := RB[7, 6];
mon_line_sn := Line.Sn; mon_line_job := RJ[8]; mon_line_alarm := Line.Alarm; mon_line_seg := Seg[8]; mon_line_n := Nst[8];
mon_line_b1 := RB[8, 1]; mon_line_b2 := RB[8, 2]; mon_line_b3 := RB[8, 3]; mon_line_b4 := RB[8, 4]; mon_line_b5 := RB[8, 5]; mon_line_b6 := RB[8, 6];
END_PROGRAM
